(* CODESYS project Simulation_Roboter.project

Project tree, tasks and I/O mapping:
  Device : CODESYS Virtual Control for Linux SL, CODESYS, order no. 2302000005, version 4.22.0.0
    application Application
      libraries: Standard, 3.5.22.0 (System); VisuDialogs, * (System); Unit Conversion Interfaces, * (Intern); CAA Mathematics, * (CAA Technical Workgroup); SM3_Math, * (CODESYS); SysProcess, * (System); CmpBitmapPool, * (System); SysProcess Implementation, * (System)
      task MainTask (cyclic, interval t#20ms, priority 1) calls MAIN_PRG
      task SoftMotion_PlanningTask (cyclic, interval t#2ms, priority 15) calls nothing
      global variables GVL_OPCUA
      visualisation Topics_Vis
      Structs/
        ST_RobotStatus/
          data type ST_RobotStatus
        ST_RobotAction/
          data type ST_RobotAction
          data type Error_Codes_RobotAction
        ST_RobotCommand/
          data type ST_RobotCommand
          data type Status_Codes_RobotCommand
        ST_Orientierung/
          data type ST_euler
          data type ST_quaternions
        ST_Roboter/
          data type ST_Pose_Axis
          data type ST_Pose_TCP
      program MAIN_PRG [FBD]
      FB_Generell/
        function block FB_MoveAction [ST]: MoveToHome, Ex1_ompl_tcp, Ex2_ompl_joint, Ex3_pilz_tcp_ptp, Ex_4_pilz_tcp_lin
        function block FB_Modes [FBD]
        function block FB_RobotStatus [ST]
        function block FB_RobotCommand [ST]
        function block FB_Watchdog [ST]
      program Ablaufkette [SFC]: Ablauf_HomePos, Ablauf_Pos1, Ablauf_Pos2, Ablauf_Pos3, Ablauf_Pos4, Ablauf_Pos5
      Funktionen/
        function FUNC_quat_to_euler [ST]
        function block FB_Quat_to_ZYZ [FBD]
        function block FB_ZYZ_to_Quat [FBD]
        function block FB_Quat_to_ZYX [FBD]
      Symbols
      image pool ImagePool
      visualisation VISU_Auto
      visualisation VISU_Startseite
      visualisation VISU_Manuell
      visualisation VISU_Konfig
      visualisation VISU_Schrittkette
  libraries: SM3_Robotics, * (CODESYS); VisuSymbols, 4.5.0.0 (System)
  text list GlobalTextList
  5ce3da45-db07-42e7-a21c-a00fff4ed8f6|C:\Users\koerp\Documents\Uni\WS2627\04_Projektarbeit-Seitz\Draw_IO\OPC_Strukut.png
  5ce3da45-db07-42e7-a21c-a00fff4ed8f6|C:\Users\koerp\Documents\Uni\WS2627\04_Projektarbeit-Seitz\Draw IO Diagramme\Screenshots\myCobotbeschriftet.png
*)

// Device/Application/Structs/ST_RobotStatus/ST_RobotStatus
// Status Client: Schnittstelle ROS2 <-> SPS
// Ist Zustand des Roboters
TYPE ST_RobotStatus :
STRUCT
	//Ist Gelenkwinkel [rad]
	Ist_Pos_Axis : ST_Pose_Axis; 	
	
	// Ist TCP Pose bezogen auf Roboterbasis
	Ist_Pos_TCP : ST_Pose_TCP;	

	//Verbindungsüberwachung mit Watchdog 
	client_connected : BOOL;
	watchdog_counter : INT;		// Überprüft serverseitige client verbindung
END_STRUCT
END_TYPE

// Device/Application/Structs/ST_RobotCommand/ST_RobotCommand
// Command Client: Schnittstelle ROS2 <-> SPS
// Manuelle Steuerung des Roboters mit MoveIt Servo
TYPE ST_RobotCommand :
STRUCT
	// Gelenke einzeln verfahren
	Mode_Axis: BOOL;					// True: Gelenk Joggen möglich
	Soll_Axis_Servo : ST_Pose_Axis;		//Richtungsvorgabe je Gelenk
	Soll_Axis_Velocity: LREAL;			// Geschwindikeitsvorgabe je Gelenk
	
	// TCP manuell verfahren 
	Mode_TCP: BOOL;						// True: Achsen Joggen möglich
	Soll_TCP_Servo : ST_Pose_TCP;		// Hinweis: Rotation wird nur mit x,y,z übergeben und nicht als Quaternion!
	Soll_TCP_Velocity: LREAL;			// Geschwindkeitsvorgabe für Verfahren
	
	//enable: zum starten und stopen des services servo_node/start_servo und stop_servo
	enable : BOOL;
	
	//Status Code mit Status Codes
	Status_Code: SINT;
	
	// Verbindungsüberwachung mit Watchdog
	client_connected: BOOL;
	watchdog_counter: INT;
END_STRUCT
END_TYPE

// Device/Application/Structs/ST_RobotAction/ST_RobotAction
TYPE ST_RobotAction :
STRUCT
	// Ausführung
	Execute : BOOL;						// TRUE-Puls 
	Error_Code : DINT;					// Ergebnis (int32 MoveItErrorCodes), 1 = SUCCESS,
										// Bedeutung siehe Error_Codes_RobotAction

	// Planer-Auswahl
	Motion_Type : STRING;				// (string pipeline_id) 'ompl' oder 'pilz_industrial_motion_planner'
	Planner_ID : STRING;				// (string planner_id) '' (leer für OMPL), 'PTP' oder 'LIN' für Pilz

	// Art des Ziels (genau eins TRUE)
	Joint_Goal : BOOL;					// TRUE: Gelenkziel -> Soll_Pos_Axis
	TCP_GOAL : BOOL;					// TRUE: kartesisches TCP-Ziel -> Soll_Pos_TCP

	// Planer-Parameter
	num_planning_attempts : DINT;		// (int32 num_planning_attempts) Anzahl Planungsversuche
	allowed_planning_time : LREAL;		// (float64 allowed_planning_time) max. Planungszeit [s]
	max_velocity_scaling : LREAL;		// (float64 max_velocity_scaling_factor) 0..1
	max_acceleration_scaling : LREAL;	// (float64 max_acceleration_scaling_factor) 0..1

	// Zieltoleranzen
	position_tolerance : LREAL;			// (float64) Toleranz TCP-Position [m], gleich für x, y, z
	orientation_tolerance : LREAL;		// (float64) Toleranz TCP-Orientierung [rad], gleich für alle Achsen
	joint_tolerance : LREAL;			// (float64) Toleranz je Gelenk [rad]

	// Zielpose Gelenke [rad]
	Soll_Pos_Axis : ST_Pose_Axis;

	// Zielpose TCP: Position [m], Orientierung als Quaternion
	Soll_Pos_TCP : ST_Pose_TCP;

	// Verbindungsüberwachung mit Watchdog
	client_connected : BOOL;		
	watchdog_counter : INT;				
END_STRUCT
END_TYPE

// Device/Application/Structs/ST_Roboter/ST_Pose_Axis
TYPE ST_Pose_Axis :
STRUCT
	// Gelenkwinkel in rad
	axis_0 : LREAL;
	axis_1 : LREAL;
	axis_2 : LREAL;
	axis_3 : LREAL;
	axis_4 : LREAL;
	axis_5 : LREAL;
END_STRUCT
END_TYPE

// Device/Application/Structs/ST_Roboter/ST_Pose_TCP
TYPE ST_Pose_TCP :
STRUCT
	// Position in m
	trans_x : LREAL;	
	trans_y :  LREAL;
	trans_z : LREAL;
	// Orientierung als Quaternion
	rot_x : LREAL;	// Imaginärteil 	
	rot_y : LREAL;	// Imaginärteil 	
	rot_z : LREAL;	// Imaginärteil 	
	rot_w : LREAL;	//Realteil
END_STRUCT
END_TYPE

// Device/Application/Structs/ST_RobotAction/Error_Codes_RobotAction
{attribute 'qualified_only'}
//{attribute 'strict'}	//CODESYS erlaubt keine TYP Umwandlungen wenn strict aktiv!
{attribute 'to_string'}

TYPE Error_Codes_RobotAction :
(
	NOT_DEFINED := 0,
    SUCCESS := 1,
    FAILURE := 99999,
    PLANNING_FAILED := -1,
    INVALID_MOTION_PLAN := -2,
    MOTION_PLAN_INVALIDATED_BY_ENVIRONMENT_CHANGE := -3,
    CONTROL_FAILED := -4,
    UNABLE_TO_AQUIRE_SENSOR_DATA := -5,
    TIMED_OUT := -6,
    PREEMPTED := -7,
    START_STATE_IN_COLLISION := -10,
    START_STATE_VIOLATES_PATH_CONSTRAINTS := -11,
    START_STATE_INVALID := -26,
    GOAL_IN_COLLISION := -12,
    GOAL_VIOLATES_PATH_CONSTRAINTS := -13,
    GOAL_CONSTRAINTS_VIOLATED := -14,
    GOAL_STATE_INVALID := -27,
    UNRECOGNIZED_GOAL_TYPE := -28,
    INVALID_GROUP_NAME := -15,
    INVALID_GOAL_CONSTRAINTS := -16,
    INVALID_ROBOT_STATE := -17,
    INVALID_LINK_NAME := -18,
    INVALID_OBJECT_NAME := -19,
    FRAME_TRANSFORM_FAILURE := -21,
    COLLISION_CHECKING_UNAVAILABLE := -22,
    ROBOT_STATE_STALE := -23,
    SENSOR_INFO_STALE := -24,
    COMMUNICATION_FAILURE := -25,
    CRASH := -29,
    ABORT := -30,
    NO_IK_SOLUTION := -31
) DINT := NOT_DEFINED;	//Standardwert
END_TYPE

// Device/Application/Structs/ST_Orientierung/ST_euler
//Eulerwinkel intrinsich ZYZ
//ZYZ intrinsisch: bezug auf mitbewegendes Koordinatensystem
//ZYZ extrinsisch: bezug auf festes Koordinatensystem
TYPE ST_euler :
STRUCT
	A : LREAL;	//Z	
	B : LREAL;	//Y
	C : LREAL;	//Z
END_STRUCT
END_TYPE

// Device/Application/Structs/ST_Orientierung/ST_quaternions
TYPE ST_quaternions :
STRUCT
	qx: LREAL;
	qy: LREAL;
	qz: LREAL;
	qw: LREAL;
END_STRUCT
END_TYPE

// Device/Application/Structs/ST_RobotCommand/Status_Codes_RobotCommand
{attribute 'qualified_only'}
//{attribute 'strict'}	//CODESYS erlaubt keine TYP Umwandlungen wenn strict aktiv!
{attribute 'to_string'}
TYPE Status_Codes_RobotCommand :
(
	SERVO_AUS := 99, //wenn Roboter nicht verbunden
	INVALID := -1,
	NO_WARNING := 0,
	DECELERATE_FOR_APPROACHING_SINGULARITY := 1,
	HALT_FOR_SINGULARITY := 2,
	DECELERATE_FOR_LEAVING_SINGULARITY := 3,
	DECELERATE_FOR_COLLISION := 4,
	HALT_FOR_COLLISION := 5,
	JOINT_BOUND := 6	// Achse hat Limit erreich
) SINT := SERVO_AUS;	//Standardwert
END_TYPE

// Device/Application/GVL_OPCUA
{attribute 'qualified_only'}
VAR_GLOBAL
// 	================ Schnittstelle OPC UA =======================================================
	// Schnittstelle Client: ROS2 <-> SPS
	RobotAction: ST_RobotAction;	// Action Client: (Bahnplannung mit MoveIt2)
	RobotStatus : ST_RobotStatus;	// Status Client: Sensorinformationen über Stand des Roboters
	RobotCommand : ST_RobotCommand;	// Command Client: /(Manuelle Steuerung mit MoveIt Servo) 
	// Schnittstelle für SoftKeys 
	// Werden von entrypoint.py Client gelesen, der dann ros2 launch Befehle startet
	Start_RViz2 : BOOL;			//Start RViz2
	Stop_RViz2: BOOL;			//Stop RViz2
	Start_OPCClients: BOOL;		//Start OPC Clients
	Stop_OPC_Clients: BOOL;		//Stop OPC Clients
	
// ================ INTERN ===================================================================	
	Execute : BOOL := FALSE;	//Taster Visu: Ausführen des MoveIt2 Befehls (Auto)
	
	// Ablaufkette
	TIPP : BOOL; 				// Zum Weiterschalten
	Start_Ablaufkette: BOOL;	// Startet Ablaufkette
	Reset_Ablaufkette: BOOL;	//setzt Schrittkette zurück
	
	Joint_Goal : BOOL;			// True: Gelenkziel vorgeben
	TCP_GOAL: BOOL;				// True: Karteisisches TCP Ziel vorgeben
	
	// TCP Sollpositionen (beuogen auf Roboterbasis)
	trans_x : LREAL;	// [m]
	trans_y : LREAL;	// [m]
	trans_z : LREAL;	// [m]
	rot_A : LREAL;		// [°]
	rot_B: LREAL;		// [°]
	rot_C: LREAL;		// [°]
	// Gelenkwinkel Sollpositionen in rad
	axis_0 : LREAL;		// [rad]
	axis_1 : LREAL;		// [rad]
	axis_2 : LREAL;		// [rad]
	axis_3 : LREAL;		// [rad]
	axis_4 : LREAL;		// [rad]
	axis_5 : LREAL;		// [rad]
	// Zieltoleranzen
	position_tolerance : LREAL;			// Toleranz TCP Position [m]
	orientation_tolerance : LREAL;		// Toleranz TCP Orientierung [rad]
	joint_tolerance: LREAL;				// Tolerant Achswinkel in [rad]

	Motion_Type : STRING;				// pipeline_id: "ompl" oder "pilz_industrial_motion_planner"
	Planner_ID : STRING;				// planner_id: " " (leer für OMPL) "PTP" oder "LIN" für Pilz

	num_planning_attempts : DINT;		// Anzahl Plannungsversuche
	allowed_planning_time : LREAL;		// max Plannungszeit in s
	max_velocity_scaling : LREAL;		// 0 .. 1 Skalierung maximale Gelenkgeschwindigkeit
	max_acceleration_scaling : LREAL;	// 0 ...1 Skalierung maximale Gelenkbeschleunigung
END_VAR

VAR_GLOBAL CONSTANT
	PI : REAL := 3.14159;
END_VAR

// Device/Application/MAIN_PRG
PROGRAM MAIN_PRG
VAR
// ======== Betriebsart ==============================================================
	Modes : FB_Modes;						// Auswahl Hand / Automatik (Hand hat Vorrang)
	
// ========Automatik ==============================================================
	// Automatik: Bewegungsauftrag an MoveIt 2 (Action Client)
	RobotAction : FB_MoveAction;			// Übergibt Sollwerte aus GVL_OPCUA an RobotAction
	trig : R_TRIG;							// Flanke von GVL_OPCUA.Execute 
	Action_zyz_to_quat : FB_ZYZ_to_Quat;	// Soll-Orientierung ZYZ -> Quaternion
	Status_Error_Codes_Action : Error_Codes_RobotAction;	// Ergebnis der Bewegung 

	// Vorgefertigte Beispielbewegungen 
	xMoveHome : BOOL;						
	xEx1_ompl_tcp : BOOL;				
	xEx2_ompl_joint : BOOL;				
	xEx3_pilz_tcp_ptp : BOOL;			
	xEx4_pilz_tcp_lin : BOOL;			

// ============Handbetrieb ==========================================================
	// Handbetrieb: Joggen über MoveIt Servo (Command Client)

	RobotCommand : FB_RobotCommand;		
	Status_Servo : Status_Codes_RobotCommand;	// Statuscode MoveIt Servo 

// ==============Istwerte========================================================
	// Istwerte und Verbindungsüberwachung (Status Client)
	RobotStatus : FB_RobotStatus;			// Watchdog Status Client
	Status_Quat_to_ZYZ : FB_Quat_to_ZYZ;	// Ist-Orientierung TCP Quaternion -> ZYZ 
END_VAR

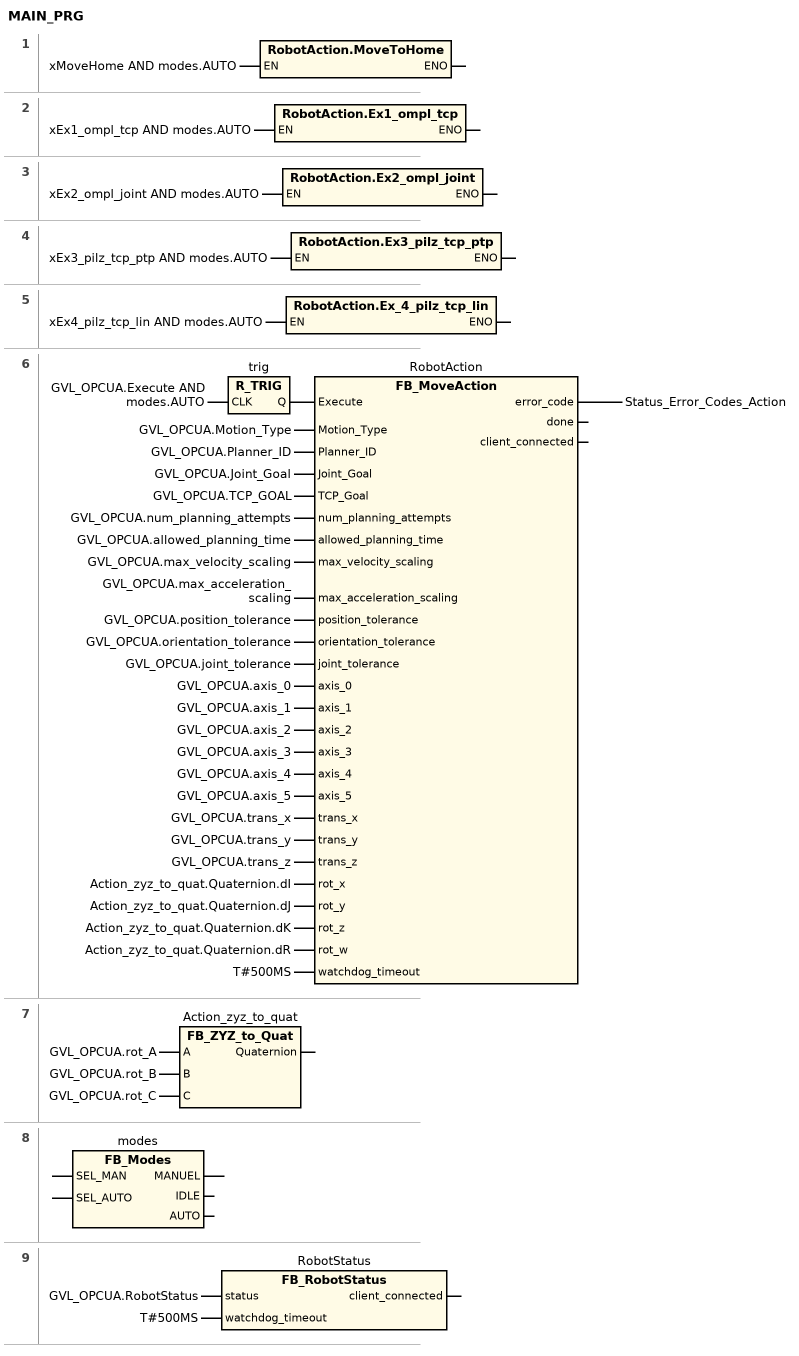
// NETWORK 1
IF xMoveHome AND modes.AUTO THEN RobotAction.MoveToHome(); END_IF

// NETWORK 2
IF xEx1_ompl_tcp AND modes.AUTO THEN RobotAction.Ex1_ompl_tcp(); END_IF

// NETWORK 3
IF xEx2_ompl_joint AND modes.AUTO THEN RobotAction.Ex2_ompl_joint(); END_IF

// NETWORK 4
IF xEx3_pilz_tcp_ptp AND modes.AUTO THEN RobotAction.Ex3_pilz_tcp_ptp(); END_IF

// NETWORK 5
IF xEx4_pilz_tcp_lin AND modes.AUTO THEN RobotAction.Ex_4_pilz_tcp_lin(); END_IF

// NETWORK 6
trig(CLK := GVL_OPCUA.Execute AND modes.AUTO); // R_TRIG
RobotAction(
    Execute := trig.Q,
    Motion_Type := GVL_OPCUA.Motion_Type,
    Planner_ID := GVL_OPCUA.Planner_ID,
    Joint_Goal := GVL_OPCUA.Joint_Goal,
    TCP_Goal := GVL_OPCUA.TCP_GOAL,
    num_planning_attempts := GVL_OPCUA.num_planning_attempts,
    allowed_planning_time := GVL_OPCUA.allowed_planning_time,
    max_velocity_scaling := GVL_OPCUA.max_velocity_scaling,
    max_acceleration_scaling := GVL_OPCUA.max_acceleration_scaling,
    position_tolerance := GVL_OPCUA.position_tolerance,
    orientation_tolerance := GVL_OPCUA.orientation_tolerance,
    joint_tolerance := GVL_OPCUA.joint_tolerance,
    axis_0 := GVL_OPCUA.axis_0,
    axis_1 := GVL_OPCUA.axis_1,
    axis_2 := GVL_OPCUA.axis_2,
    axis_3 := GVL_OPCUA.axis_3,
    axis_4 := GVL_OPCUA.axis_4,
    axis_5 := GVL_OPCUA.axis_5,
    trans_x := GVL_OPCUA.trans_x,
    trans_y := GVL_OPCUA.trans_y,
    trans_z := GVL_OPCUA.trans_z,
    rot_x := Action_zyz_to_quat.Quaternion.dI,
    rot_y := Action_zyz_to_quat.Quaternion.dJ,
    rot_z := Action_zyz_to_quat.Quaternion.dK,
    rot_w := Action_zyz_to_quat.Quaternion.dR,
    watchdog_timeout := T#500MS); // FB_MoveAction
Status_Error_Codes_Action := RobotAction.error_code;

// NETWORK 7
Action_zyz_to_quat(A := GVL_OPCUA.rot_A, B := GVL_OPCUA.rot_B, C := GVL_OPCUA.rot_C); // FB_ZYZ_to_Quat

// NETWORK 8
modes(); // FB_Modes

// NETWORK 9
RobotStatus(status := GVL_OPCUA.RobotStatus, watchdog_timeout := T#500MS); // FB_RobotStatus

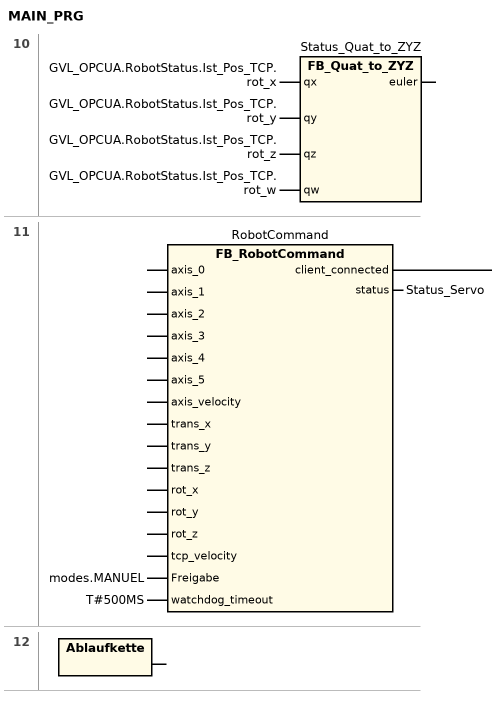
// NETWORK 10
Status_Quat_to_ZYZ(
    qx := GVL_OPCUA.RobotStatus.Ist_Pos_TCP.rot_x,
    qy := GVL_OPCUA.RobotStatus.Ist_Pos_TCP.rot_y,
    qz := GVL_OPCUA.RobotStatus.Ist_Pos_TCP.rot_z,
    qw := GVL_OPCUA.RobotStatus.Ist_Pos_TCP.rot_w); // FB_Quat_to_ZYZ

// NETWORK 11
RobotCommand(Freigabe := modes.MANUEL, watchdog_timeout := T#500MS, status => Status_Servo); // FB_RobotCommand

// NETWORK 12
Ablaufkette();

END_PROGRAM

// Device/Application/FB_Generell/FB_MoveAction
FUNCTION_BLOCK FB_MoveAction
// Übergabe von Gelenk oder ZCP Ziel an ROS2 Client
VAR_INPUT
    Execute : BOOL;

    Motion_Type : STRING;
    Planner_ID : STRING;

    Joint_Goal : BOOL;
    TCP_Goal : BOOL;

    num_planning_attempts : DINT;
    allowed_planning_time : LREAL;

    max_velocity_scaling : LREAL;
    max_acceleration_scaling : LREAL;

    position_tolerance : LREAL;
    orientation_tolerance : LREAL;
	joint_tolerance: LREAL;

    // Joints
    axis_0 : LREAL;
    axis_1 : LREAL;
    axis_2 : LREAL;
    axis_3 : LREAL;
    axis_4 : LREAL;
    axis_5 : LREAL;

    // TCP
    trans_x : LREAL;
    trans_y : LREAL;
    trans_z : LREAL;
    rot_x : LREAL;
    rot_y : LREAL;
    rot_z : LREAL;
    rot_w : LREAL;
	
	watchdog_timeout : TIME := T#500MS;	//Timeout des Watchdogs
END_VAR
VAR_OUTPUT
	error_code:DINT;
	done : BOOL;
	//Watchdog
	client_connected : BOOL;
END_VAR
VAR
	watchdog : FB_Watchdog;
END_VAR

//Watchdog aktualisieren
watchdog(watchdog_counter := GVL_OPCUA.RobotAction.watchdog_counter, timeout := watchdog_timeout);
client_connected := watchdog.client_connected;

// Execute
GVL_OPCUA.RobotAction.Execute := Execute;

// Allgemein
GVL_OPCUA.RobotAction.Motion_Type := Motion_Type;
GVL_OPCUA.RobotAction.Planner_ID := Planner_ID;

GVL_OPCUA.RobotAction.Joint_Goal := Joint_Goal;
GVL_OPCUA.RobotAction.TCP_GOAL := TCP_Goal;

GVL_OPCUA.RobotAction.num_planning_attempts := num_planning_attempts;
GVL_OPCUA.RobotAction.allowed_planning_time := allowed_planning_time;

GVL_OPCUA.RobotAction.max_velocity_scaling := max_velocity_scaling;
GVL_OPCUA.RobotAction.max_acceleration_scaling := max_acceleration_scaling;

GVL_OPCUA.RobotAction.position_tolerance := position_tolerance;
GVL_OPCUA.RobotAction.orientation_tolerance := orientation_tolerance;
GVL_OPCUA.RobotAction.joint_tolerance := joint_tolerance;

// Joints
GVL_OPCUA.RobotAction.Soll_Pos_Axis.axis_0 := axis_0;
GVL_OPCUA.RobotAction.Soll_Pos_Axis.axis_1 := axis_1;
GVL_OPCUA.RobotAction.Soll_Pos_Axis.axis_2 := axis_2;
GVL_OPCUA.RobotAction.Soll_Pos_Axis.axis_3 := axis_3;
GVL_OPCUA.RobotAction.Soll_Pos_Axis.axis_4 := axis_4;
GVL_OPCUA.RobotAction.Soll_Pos_Axis.axis_5 := axis_5;


// TCP
GVL_OPCUA.RobotAction.Soll_Pos_TCP.trans_x := trans_x;
GVL_OPCUA.RobotAction.Soll_Pos_TCP.trans_y := trans_y;
GVL_OPCUA.RobotAction.Soll_Pos_TCP.trans_z := trans_z;

GVL_OPCUA.RobotAction.Soll_Pos_TCP.rot_x := rot_x;
GVL_OPCUA.RobotAction.Soll_Pos_TCP.rot_y := rot_y;
GVL_OPCUA.RobotAction.Soll_Pos_TCP.rot_z := rot_z;
GVL_OPCUA.RobotAction.Soll_Pos_TCP.rot_w := rot_w;

//OUTPUT
error_code := GVL_OPCUA.RobotAction.Error_Code;
IF error_code = 1 THEN
	done := TRUE;
ELSE 
	done := FALSE;
END_IF

ACTION MoveToHome:
//HomePosition
GVL_OPCUA.Joint_Goal := TRUE;
GVL_OPCUA.TCP_Goal := FALSE;

GVL_OPCUA.axis_0 := 0.0;
GVL_OPCUA.axis_1 := 0.0;
GVL_OPCUA.axis_2 := 0.0;
GVL_OPCUA.axis_3 := 0.0;
GVL_OPCUA.axis_4 := 0.0;
GVL_OPCUA.axis_5 := 0.0;

GVL_OPCUA.joint_tolerance := 0.005;

GVL_OPCUA.Motion_Type := 'ompl';
GVL_OPCUA.Planner_ID := '';

GVL_OPCUA.num_planning_attempts := 5;
GVL_OPCUA.allowed_planning_time := 5;
GVL_OPCUA.max_velocity_scaling := 0.1;
GVL_OPCUA.max_acceleration_scaling := 0.1;
END_ACTION

ACTION Ex1_ompl_tcp:
GVL_OPCUA.Joint_Goal := FALSE;
GVL_OPCUA.TCP_Goal := TRUE;

GVL_OPCUA.trans_x := 0.114;
GVL_OPCUA.trans_y := -0.019;
GVL_OPCUA.trans_z := 0.357;
GVL_OPCUA.rot_A := 0.0;
GVL_OPCUA.rot_B := 90.0;
GVL_OPCUA.rot_C := -90.0;

GVL_OPCUA.position_tolerance := 0.02;
GVL_OPCUA.orientation_tolerance := 0.05;

GVL_OPCUA.Motion_Type := 'ompl';
GVL_OPCUA.Planner_ID := '';

GVL_OPCUA.num_planning_attempts := 5;
GVL_OPCUA.allowed_planning_time := 5;
GVL_OPCUA.max_velocity_scaling := 0.2;
GVL_OPCUA.max_acceleration_scaling := 0.2;
END_ACTION

ACTION Ex2_ompl_joint:
GVL_OPCUA.Joint_Goal := TRUE;
GVL_OPCUA.TCP_Goal := FALSE;

GVL_OPCUA.axis_0 := 0.1;
GVL_OPCUA.axis_1 := -1.65;
GVL_OPCUA.axis_2 := 1.7;
GVL_OPCUA.axis_3 := 0.1;
GVL_OPCUA.axis_4 := 0.2;
GVL_OPCUA.axis_5 := 0.3;

GVL_OPCUA.Motion_Type := 'ompl';
GVL_OPCUA.Planner_ID := '';

GVL_OPCUA.joint_tolerance := 0.01;

GVL_OPCUA.num_planning_attempts := 5;
GVL_OPCUA.allowed_planning_time := 5;
GVL_OPCUA.max_velocity_scaling := 0.2;
GVL_OPCUA.max_acceleration_scaling := 0.2;
END_ACTION

ACTION Ex3_pilz_tcp_ptp:
GVL_OPCUA.Joint_Goal := FALSE;
GVL_OPCUA.TCP_Goal := TRUE;

GVL_OPCUA.trans_x := 0.17;
GVL_OPCUA.trans_y := -0.04;
GVL_OPCUA.trans_z := 0.22;
GVL_OPCUA.rot_A := 0.0;
GVL_OPCUA.rot_B := 90.0;
GVL_OPCUA.rot_C := -90.0;

GVL_OPCUA.position_tolerance := 0.02;
GVL_OPCUA.orientation_tolerance := 0.05;

GVL_OPCUA.Motion_Type := 'pilz_industrial_motion_planner';
GVL_OPCUA.Planner_ID := 'PTP';

GVL_OPCUA.num_planning_attempts := 10;
GVL_OPCUA.allowed_planning_time := 10;
GVL_OPCUA.max_velocity_scaling := 0.05;
GVL_OPCUA.max_acceleration_scaling := 0.05;
END_ACTION

ACTION Ex_4_pilz_tcp_lin:
GVL_OPCUA.Joint_Goal := FALSE;
GVL_OPCUA.TCP_Goal := TRUE;

GVL_OPCUA.trans_x := 0.2;
GVL_OPCUA.trans_y := -0.041;
GVL_OPCUA.trans_z := 0.3;
GVL_OPCUA.rot_A := 0.0;
GVL_OPCUA.rot_B := 90.0;
GVL_OPCUA.rot_C := -90.0;

GVL_OPCUA.Motion_Type := 'pilz_industrial_motion_planner';
GVL_OPCUA.Planner_ID := 'LIN';

GVL_OPCUA.position_tolerance := 0.02;
GVL_OPCUA.orientation_tolerance := 0.05;

GVL_OPCUA.num_planning_attempts := 10;
GVL_OPCUA.allowed_planning_time := 10;
GVL_OPCUA.max_velocity_scaling := 0.005;
GVL_OPCUA.max_acceleration_scaling := 0.005;
END_ACTION

END_FUNCTION_BLOCK

// Device/Application/FB_Generell/FB_Watchdog
FUNCTION_BLOCK FB_Watchdog
VAR_INPUT
	Watchdog_counter: INT;	// Zähler im ROS2 Programm
	Timeout : TIME := T#500MS;
END_VAR
VAR
	//Watchdog
	Watchdog_counter_old : INT := 0;
	Timer : TON;
END_VAR
VAR_OUTPUT
	client_connected: BOOL;	//Anzeige ob verbunden
END_VAR

//Watchdog zum Testen ob noch mit Client verbunden!
IF Watchdog_counter <> Watchdog_counter_old THEN
	Watchdog_counter_old :=  Watchdog_counter;
    client_connected := TRUE;
    Timer(IN := FALSE);
ELSE
    Timer(IN := TRUE,PT := Timeout );
END_IF;
IF Timer.Q THEN
    client_connected := FALSE;
END_IF;

END_FUNCTION_BLOCK

// Device/Application/Funktionen/FB_ZYZ_to_Quat
FUNCTION_BLOCK FB_ZYZ_to_Quat
VAR_INPUT
	A : LREAL;
	B: LREAL;
	C: LREAL;
END_VAR
VAR_OUTPUT
	Quaternion: SMC_Quat;
END_VAR
VAR
	Rotation_Matrix: SMC_Matrix3;
END_VAR

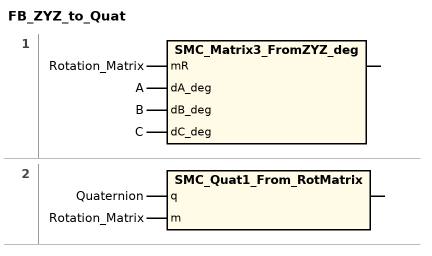
// NETWORK 1
SMC_Matrix3_FromZYZ_deg(mR := Rotation_Matrix, dA_deg := A, dB_deg := B, dC_deg := C);

// NETWORK 2
SMC_Quat1_From_RotMatrix(q := Quaternion, m := Rotation_Matrix);

END_FUNCTION_BLOCK

// Device/Application/FB_Generell/FB_Modes
FUNCTION_BLOCK FB_Modes	// Betriebsartenumschaltung mit Betriebsartenhierachie MAN > AUTO
VAR_INPUT
	SEL_MAN : BOOL;
	SEL_AUTO: BOOL;
END_VAR
VAR_OUTPUT
	MANUEL : BOOL;	//z1
	IDLE: BOOL;		//z0
	AUTO: BOOL;		//z2
END_VAR
VAR
	z0, z1, z2 : BOOL;
	H1, H2: RS;
	z: INT;
END_VAR
VAR // added by the converter: edge detectors and wires of the graphical bodies
    _w1, _w2, _w3 : BOOL;
END_VAR

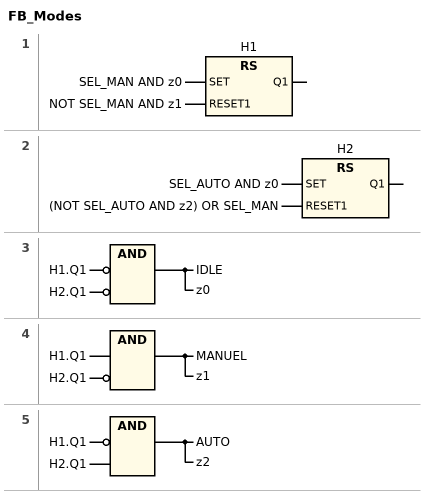
// NETWORK 1
H1(SET := SEL_MAN AND z0, RESET1 := NOT SEL_MAN AND z1); // RS

// NETWORK 2
H2(SET := SEL_AUTO AND z0, RESET1 := (NOT SEL_AUTO AND z2) OR SEL_MAN); // RS

// NETWORK 3
_w1 := NOT H1.Q1 AND NOT H2.Q1;
IDLE := _w1;
z0 := _w1;

// NETWORK 4
_w2 := H1.Q1 AND NOT H2.Q1;
MANUEL := _w2;
z1 := _w2;

// NETWORK 5
_w3 := NOT H1.Q1 AND H2.Q1;
AUTO := _w3;
z2 := _w3;

END_FUNCTION_BLOCK

// Device/Application/FB_Generell/FB_RobotStatus
FUNCTION_BLOCK FB_RobotStatus
VAR_INPUT
	status: ST_RobotStatus;
	watchdog_timeout: TIME := T#500MS;
END_VAR
VAR_OUTPUT
	client_connected : BOOL;
END_VAR
VAR
	watchdog : FB_Watchdog;
END_VAR

//Watchdog aktualisieren
watchdog(watchdog_counter := status.watchdog_counter, timeout := watchdog_timeout);
client_connected := watchdog.client_connected;

END_FUNCTION_BLOCK

// Device/Application/Funktionen/FB_Quat_to_ZYZ
FUNCTION_BLOCK FB_Quat_to_ZYZ
VAR_INPUT
	qx : LREAL;
	qy: LREAL;
	qz:LREAL;
	qw : LREAL;

END_VAR
VAR_OUTPUT
	euler : ST_euler;
END_VAR
VAR
	Quaternion: SMC_Quat;
	Rotation_Matrix: SMC_Matrix3;
END_VAR

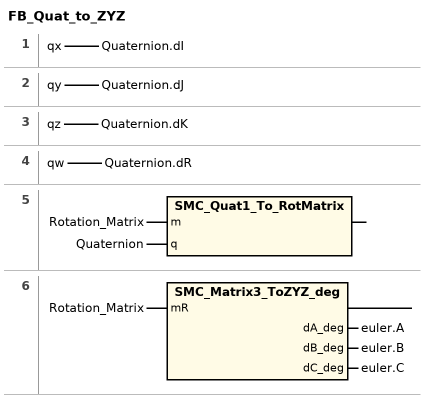
// NETWORK 1
Quaternion.dI := qx;

// NETWORK 2
Quaternion.dJ := qy;

// NETWORK 3
Quaternion.dK := qz;

// NETWORK 4
Quaternion.dR := qw;

// NETWORK 5
SMC_Quat1_To_RotMatrix(m := Rotation_Matrix, q := Quaternion);

// NETWORK 6
SMC_Matrix3_ToZYZ_deg(mR := Rotation_Matrix, dA_deg => euler.A, dB_deg => euler.B, dC_deg => euler.C);

END_FUNCTION_BLOCK

// Device/Application/FB_Generell/FB_RobotCommand
FUNCTION_BLOCK FB_RobotCommand
VAR_INPUT
	axis_0 : LREAL;
	axis_1 : LREAL;
	axis_2: LREAL;
	axis_3 : LREAL;
	axis_4 : LREAL;
	axis_5 : LREAL;
	axis_velocity : LREAL;
	
	trans_x : LREAL;
	trans_y : LREAL;
	trans_z : LREAL;
	rot_x : LREAL;
	rot_y : LREAL;
	rot_z : LREAL;
	tcp_velocity : LREAL;
	
	//Allgemein
	Freigabe:BOOL:=FALSE;
	
	watchdog_timeout: TIME := T#500MS;
END_VAR
VAR_OUTPUT
	// Watchdog
	client_connected : BOOL;
	// Status Meldung
	status: SINT;	//Datentyp INT8
END_VAR
VAR
	//Watchdog
	watchdog : FB_Watchdog;
END_VAR

//Watchdog aktualisieren
watchdog(watchdog_counter := GVL_OPCUA.RobotCommand.watchdog_counter, timeout := watchdog_timeout);
client_connected := watchdog.client_connected;

IF Freigabe THEN	//Freigabe wenn manueller Betrieb
	GVL_OPCUA.RobotCommand.Soll_Axis_Servo.axis_0 := axis_0;
	GVL_OPCUA.RobotCommand.Soll_Axis_Servo.axis_1 := axis_1;
	GVL_OPCUA.RobotCommand.Soll_Axis_Servo.axis_2 := axis_2;
	GVL_OPCUA.RobotCommand.Soll_Axis_Servo.axis_3 := axis_3;
	GVL_OPCUA.RobotCommand.Soll_Axis_Servo.axis_4 := axis_4;
	GVL_OPCUA.RobotCommand.Soll_Axis_Servo.axis_5 := axis_5;
	GVL_OPCUA.RobotCommand.Soll_Axis_Velocity := axis_velocity;
	
	GVL_OPCUA.RobotCommand.Soll_TCP_Servo.trans_x := trans_x;
	GVL_OPCUA.RobotCommand.Soll_TCP_Servo.trans_y := trans_y;
	GVL_OPCUA.RobotCommand.Soll_TCP_Servo.trans_z := trans_z;
	GVL_OPCUA.RobotCommand.Soll_TCP_Servo.rot_x := rot_x;
	GVL_OPCUA.RobotCommand.Soll_TCP_Servo.rot_y := rot_y;
	GVL_OPCUA.RobotCommand.Soll_TCP_Servo.rot_z := rot_z;
	GVL_OPCUA.RobotCommand.Soll_TCP_Velocity := tcp_velocity;
	
	// start der /servo_node/start_servo
	GVL_OPCUA.RobotCommand.enable := TRUE;
	
ELSE
	GVL_OPCUA.RobotCommand.enable := FALSE;
END_IF

// Status Code
status := GVL_OPCUA.RobotCommand.Status_Code;

END_FUNCTION_BLOCK

// Device/Application/Ablaufkette
PROGRAM Ablaufkette
VAR
	SFCCurrentStep : STRING;
END_VAR

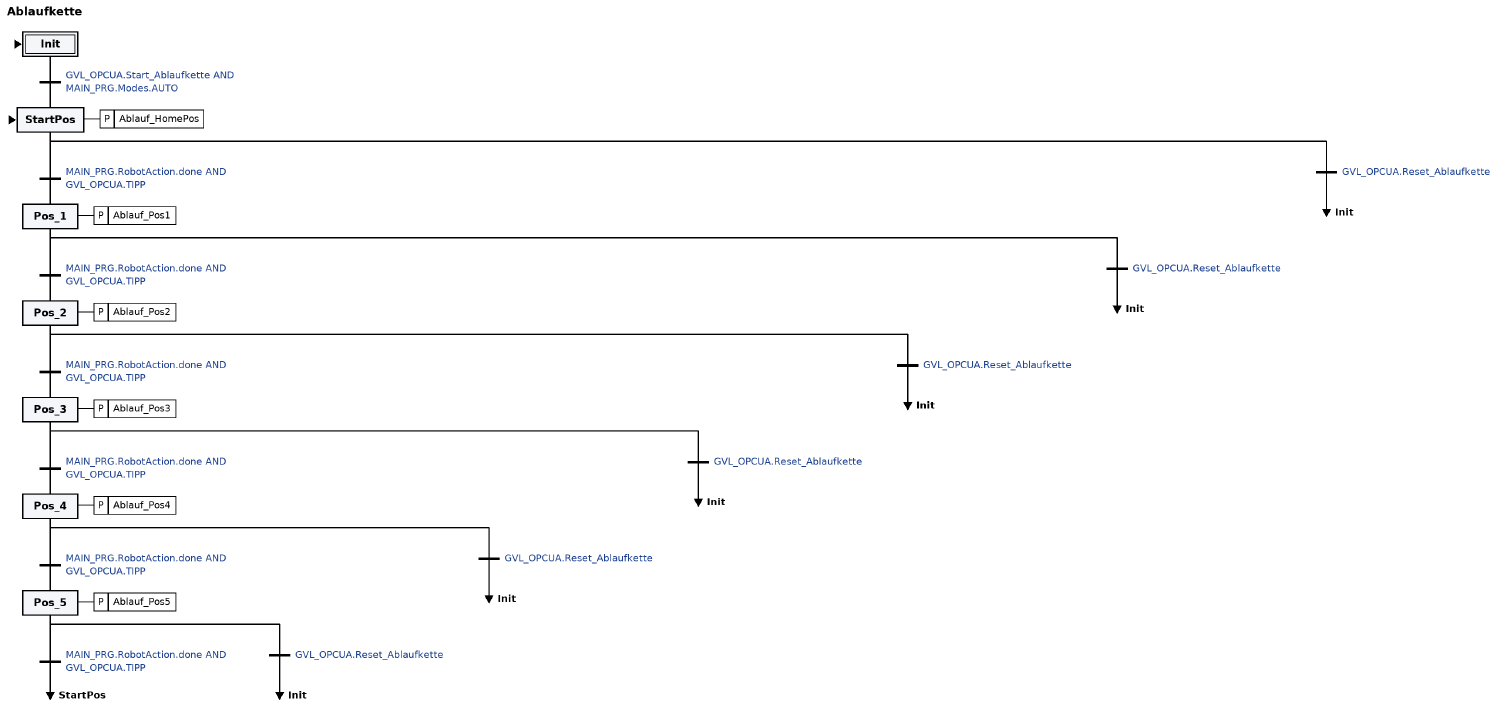
INITIAL_STEP Init:
END_STEP
TRANSITION FROM Init TO StartPos
    := GVL_OPCUA.Start_Ablaufkette AND MAIN_PRG.Modes.AUTO;
END_TRANSITION
STEP StartPos:  // min time t#1s
    Ablauf_HomePos(P);
END_STEP
TRANSITION FROM StartPos TO Pos_1
    := MAIN_PRG.RobotAction.done AND GVL_OPCUA.TIPP;
END_TRANSITION
TRANSITION FROM StartPos TO Init
    := GVL_OPCUA.Reset_Ablaufkette;
END_TRANSITION
STEP Pos_1:  // min time t#1s
    Ablauf_Pos1(P);
END_STEP
TRANSITION FROM Pos_1 TO Pos_2
    := MAIN_PRG.RobotAction.done AND GVL_OPCUA.TIPP;
END_TRANSITION
TRANSITION FROM Pos_1 TO Init
    := GVL_OPCUA.Reset_Ablaufkette;
END_TRANSITION
STEP Pos_2:  // min time t#1s
    Ablauf_Pos2(P);
END_STEP
TRANSITION FROM Pos_2 TO Pos_3
    := MAIN_PRG.RobotAction.done AND GVL_OPCUA.TIPP;
END_TRANSITION
TRANSITION FROM Pos_2 TO Init
    := GVL_OPCUA.Reset_Ablaufkette;
END_TRANSITION
STEP Pos_3:  // min time t#1s
    Ablauf_Pos3(P);
END_STEP
TRANSITION FROM Pos_3 TO Pos_4
    := MAIN_PRG.RobotAction.done AND GVL_OPCUA.TIPP;
END_TRANSITION
TRANSITION FROM Pos_3 TO Init
    := GVL_OPCUA.Reset_Ablaufkette;
END_TRANSITION
STEP Pos_4:  // min time t#1s
    Ablauf_Pos4(P);
END_STEP
TRANSITION FROM Pos_4 TO Pos_5
    := MAIN_PRG.RobotAction.done AND GVL_OPCUA.TIPP;
END_TRANSITION
TRANSITION FROM Pos_4 TO Init
    := GVL_OPCUA.Reset_Ablaufkette;
END_TRANSITION
STEP Pos_5:  // min time t#1s
    Ablauf_Pos5(P);
END_STEP
TRANSITION FROM Pos_5 TO StartPos
    := MAIN_PRG.RobotAction.done AND GVL_OPCUA.TIPP;
END_TRANSITION
TRANSITION FROM Pos_5 TO Init
    := GVL_OPCUA.Reset_Ablaufkette;
END_TRANSITION

ACTION Ablauf_HomePos:
GVL_OPCUA.Joint_Goal := TRUE;
GVL_OPCUA.TCP_Goal := FALSE;

GVL_OPCUA.axis_0 := 0.10;
GVL_OPCUA.axis_1 := -0.1;
GVL_OPCUA.axis_2 := -1.6;
GVL_OPCUA.axis_3 := 1.7;
GVL_OPCUA.axis_4 := 0.1;
GVL_OPCUA.axis_5 := 0.2;

GVL_OPCUA.joint_tolerance := 0.01;

GVL_OPCUA.Motion_Type := 'ompl';
GVL_OPCUA.Planner_ID := '';

GVL_OPCUA.num_planning_attempts := 10;
GVL_OPCUA.allowed_planning_time := 10;

GVL_OPCUA.max_velocity_scaling := 0.2;
GVL_OPCUA.max_acceleration_scaling := 0.2;
END_ACTION

ACTION Ablauf_Pos1:
GVL_OPCUA.Joint_Goal := FALSE;
GVL_OPCUA.TCP_Goal := TRUE;

GVL_OPCUA.trans_x := 0.18;
GVL_OPCUA.trans_y := -0.0;
GVL_OPCUA.trans_z := 0.3;

GVL_OPCUA.rot_A := 0.0;
GVL_OPCUA.rot_B := 90.0;
GVL_OPCUA.rot_C := -90.0;

GVL_OPCUA.position_tolerance := 0.005;
GVL_OPCUA.orientation_tolerance := 0.05;

GVL_OPCUA.Motion_Type := 'ompl';
GVL_OPCUA.Planner_ID := '';

GVL_OPCUA.num_planning_attempts := 10;
GVL_OPCUA.allowed_planning_time := 10;
GVL_OPCUA.max_velocity_scaling := 0.1;
GVL_OPCUA.max_acceleration_scaling := 0.1;
END_ACTION

ACTION Ablauf_Pos2:
GVL_OPCUA.Joint_Goal := FALSE;
GVL_OPCUA.TCP_Goal := TRUE;

GVL_OPCUA.trans_x := 0.18;
GVL_OPCUA.trans_y := 0.05;
GVL_OPCUA.trans_z := 0.3;

GVL_OPCUA.rot_A := 0.0;
GVL_OPCUA.rot_B := 90.0;
GVL_OPCUA.rot_C := -90.0;

GVL_OPCUA.position_tolerance := 0.005;
GVL_OPCUA.orientation_tolerance := 0.05;

GVL_OPCUA.Motion_Type := 'pilz_industrial_motion_planner';
GVL_OPCUA.Planner_ID := 'PTP';

GVL_OPCUA.num_planning_attempts := 10;
GVL_OPCUA.allowed_planning_time := 10;
GVL_OPCUA.max_velocity_scaling := 0.1;
GVL_OPCUA.max_acceleration_scaling := 0.1;
END_ACTION

ACTION Ablauf_Pos3:
GVL_OPCUA.Joint_Goal := FALSE;
GVL_OPCUA.TCP_Goal := TRUE;

GVL_OPCUA.trans_x := 0.18;
GVL_OPCUA.trans_y := 0.05;
GVL_OPCUA.trans_z := 0.2;

GVL_OPCUA.rot_A := 0.0;
GVL_OPCUA.rot_B := 90.0;
GVL_OPCUA.rot_C := -90.0;

GVL_OPCUA.position_tolerance := 0.005;
GVL_OPCUA.orientation_tolerance := 0.05;

GVL_OPCUA.Motion_Type := 'pilz_industrial_motion_planner';
GVL_OPCUA.Planner_ID := 'PTP';

GVL_OPCUA.num_planning_attempts := 10;
GVL_OPCUA.allowed_planning_time := 10;
GVL_OPCUA.max_velocity_scaling := 0.1;
GVL_OPCUA.max_acceleration_scaling := 0.1;
END_ACTION

ACTION Ablauf_Pos4:
GVL_OPCUA.Joint_Goal := FALSE;
GVL_OPCUA.TCP_Goal := TRUE;

GVL_OPCUA.trans_x := 0.18;
GVL_OPCUA.trans_y := -0.05;
GVL_OPCUA.trans_z := 0.2;

GVL_OPCUA.rot_A := 0.0;
GVL_OPCUA.rot_B := 90.0;
GVL_OPCUA.rot_C := -90.0;

GVL_OPCUA.position_tolerance := 0.005;
GVL_OPCUA.orientation_tolerance := 0.05;

GVL_OPCUA.Motion_Type := 'pilz_industrial_motion_planner';
GVL_OPCUA.Planner_ID := 'PTP';

GVL_OPCUA.num_planning_attempts := 10;
GVL_OPCUA.allowed_planning_time := 10;
GVL_OPCUA.max_velocity_scaling := 0.1;
GVL_OPCUA.max_acceleration_scaling := 0.1;
END_ACTION

ACTION Ablauf_Pos5:
GVL_OPCUA.Joint_Goal := FALSE;
GVL_OPCUA.TCP_Goal := TRUE;

GVL_OPCUA.trans_x := 0.18;
GVL_OPCUA.trans_y := -0.05;
GVL_OPCUA.trans_z := 0.3;

GVL_OPCUA.rot_A := 0.0;
GVL_OPCUA.rot_B := 90.0;
GVL_OPCUA.rot_C := -90.0;

GVL_OPCUA.position_tolerance := 0.005;
GVL_OPCUA.orientation_tolerance := 0.05;

GVL_OPCUA.Motion_Type := 'pilz_industrial_motion_planner';
GVL_OPCUA.Planner_ID := 'PTP';

GVL_OPCUA.num_planning_attempts := 10;
GVL_OPCUA.allowed_planning_time := 10;
GVL_OPCUA.max_velocity_scaling := 0.1;
GVL_OPCUA.max_acceleration_scaling := 0.1;
END_ACTION

END_PROGRAM

// Device/Application/Funktionen/FUNC_quat_to_euler
FUNCTION FUNC_quat_to_euler : ST_euler
VAR_INPUT
	qx : LREAL;
	qy : LREAL;
	qz : LREAL;
	qw : LREAL;
END_VAR
VAR
	r11, r12, r13, r21, r22, r23, r31, r32, r33 : LREAL;
	const_epsilon : LREAL := 1.0E-6; // Toleranz für Gimbal Lock
	result : ST_euler;
	
END_VAR

//Quaternion -> Euler mit ZYZ (intrinsisch) 
//Ausgabe der Euler Winkel in Grad
//Rotationsmatrix Quaternion
r11 := 1.0 - 2.0 * (qy*qy + qz*qz);
r12 := 2.0 * (qx*qy - qz*qw);
r13 := 2.0 * (qx*qz + qy*qw);

r21 := 2.0 * (qx*qy + qz*qw);
r22 := 1.0 - 2.0 * (qx*qx + qz*qz);
r23 := 2.0 * (qy*qz - qx*qw);

r31 := 2.0 * (qx*qz - qy*qw);
r32 := 2.0 * (qy*qz + qx*qw);
r33 := 1.0 - 2.0 * (qx*qx + qy*qy);

result.B := MATH.atan2_func(SQRT(r31*r31+r32*r32),r33);

IF result.B < const_epsilon THEN
	//Gimbal Lock Nordpol
	result.A := 0.0;
	result.C := MATH.atan2_func(r21,r11);
	
ELSIF result.B > (MATH.PI - const_epsilon) THEN
	//Gimbal Lock Südpol
	result.A := 0.0;
	result.C := MATH.atan2_func(-r21,-r11);
ELSE
	//normal
	result.A := MATH.atan2_func(r23,r13);
	result.C := MATH.atan2_func(r32,-r31);
	
END_IF

result.A := result.A * (180.0/MATH.PI);
result.B := result.B * (180.0/MATH.PI);
result.C := result.C * (180.0/MATH.PI);

FUNC_quat_to_euler := result;

END_FUNCTION

// Device/Application/Funktionen/FB_Quat_to_ZYX
FUNCTION_BLOCK FB_Quat_to_ZYX
VAR_INPUT
	qx : LREAL;
	qy: LREAL;
	qz:LREAL;
	qw : LREAL;

END_VAR
VAR_OUTPUT
	euler : ST_euler;
END_VAR
VAR
	Quaternion: SMC_Quat;
	Rotation_Matrix: SMC_Matrix3;
END_VAR

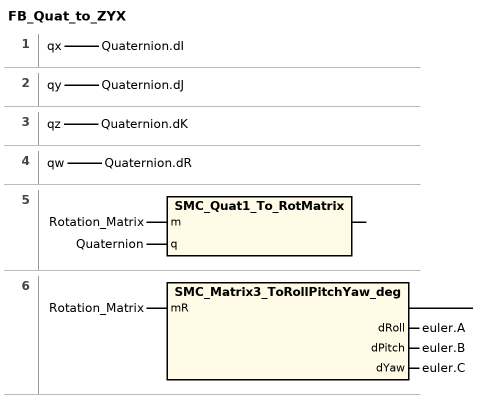
// NETWORK 1
Quaternion.dI := qx;

// NETWORK 2
Quaternion.dJ := qy;

// NETWORK 3
Quaternion.dK := qz;

// NETWORK 4
Quaternion.dR := qw;

// NETWORK 5
SMC_Quat1_To_RotMatrix(m := Rotation_Matrix, q := Quaternion);

// NETWORK 6
SMC_Matrix3_ToRollPitchYaw_deg(mR := Rotation_Matrix, dRoll => euler.A, dPitch => euler.B, dYaw => euler.C);

END_FUNCTION_BLOCK

// Device/Application/Topics_Vis
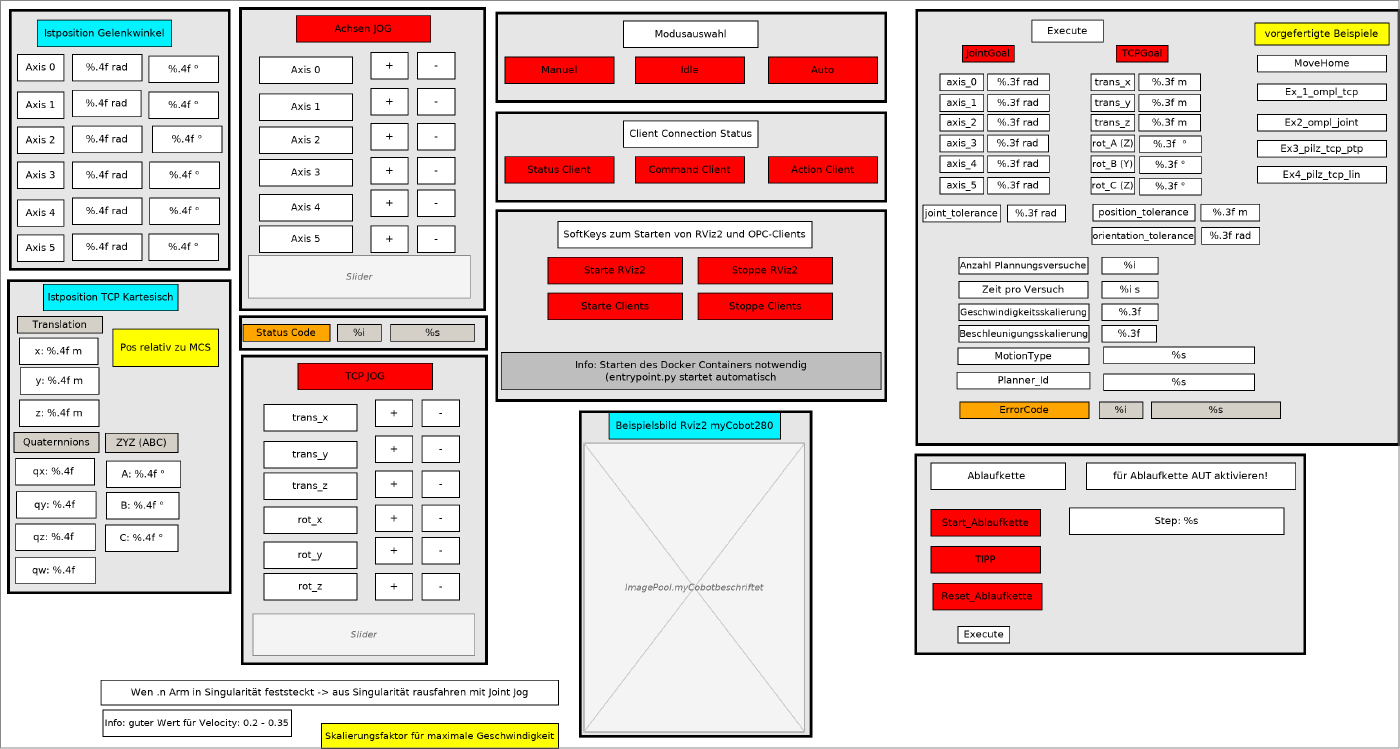
VISUALIZATION Topics_Vis  // 1557x834
    Rectangle (266,351 276x39)
    Rectangle (266,8 274x338)
    Rectangle (644,457 259x364)
    Rectangle (551,233 435x214)
    Rectangle (8,311 249x350)
    Rectangle (1018,10 539x486)
    Rectangle (551,13 435x101)
    Rectangle (10,10 246x291)
    Rectangle (41,22 150x30), "Istposition Gelenkwinkel"
    Rectangle (48,316 150x30), "Istposition TCP Kartesisch"
    Rectangle (21,376 88x30), "x: %.4f m", text variable: MAIN_PRG.RobotStatus.tcp_pose.trans_x
    Rectangle (22,409 88x30), "y: %.4f m", text variable: MAIN_PRG.RobotStatus.tcp_pose.trans_y
    Rectangle (21,445 89x30), "z: %.4f m", text variable: MAIN_PRG.RobotStatus.tcp_pose.trans_z
    Rectangle (17,510 88x30), "qx: %.4f", text variable: MAIN_PRG.RobotStatus.tcp_pose.rot_x
    Rectangle (18,547 89x30), "qy: %.4f", text variable: MAIN_PRG.RobotStatus.tcp_pose.rot_y
    Rectangle (17,583 89x30), "qz: %.4f", text variable: MAIN_PRG.RobotStatus.tcp_pose.rot_z
    Rectangle (17,620 89x30), "qw: %.4f", text variable: MAIN_PRG.RobotStatus.tcp_pose.rot_w
    Rectangle (412,58 42x30), "+"
        OnMouseDown: execute { MAIN_PRG.RobotCommand.axis_0 := +1; }
        OnMouseUp: execute { MAIN_PRG.RobotCommand.axis_0 := 0; }
    Rectangle (464,58 42x30), "-"
        OnMouseDown: execute { MAIN_PRG.RobotCommand.axis_0 := -1; }
        OnMouseUp: execute { MAIN_PRG.RobotCommand.axis_0 := 0; }
    Rectangle (412,98 42x30), "+"
        OnMouseDown: execute { MAIN_PRG.RobotCommand.axis_1 := +1; }
        OnMouseUp: execute { MAIN_PRG.RobotCommand.axis_1 := 0; }
    Rectangle (464,137 42x30), "-"
        OnMouseDown: execute { MAIN_PRG.RobotCommand.axis_2 := -1; }
        OnMouseUp: execute { MAIN_PRG.RobotCommand.axis_2 := 0; }
    Rectangle (412,137 42x30), "+"
        OnMouseDown: execute { MAIN_PRG.RobotCommand.axis_2 := +1; }
        OnMouseUp: execute { MAIN_PRG.RobotCommand.axis_2 := 0; }
    Rectangle (412,175 42x30), "+"
        OnMouseDown: execute { MAIN_PRG.RobotCommand.axis_3 := +1; }
        OnMouseUp: execute { MAIN_PRG.RobotCommand.axis_3 := 0; }
    Rectangle (464,98 42x30), "-"
        OnMouseDown: execute { MAIN_PRG.RobotCommand.axis_1 := -1; }
        OnMouseUp: execute { MAIN_PRG.RobotCommand.axis_1 := 0; }
    Rectangle (464,175 42x30), "-"
        OnMouseDown: execute { MAIN_PRG.RobotCommand.axis_3 := -1; }
        OnMouseUp: execute { MAIN_PRG.RobotCommand.axis_3 := 0; }
    Rectangle (412,211 42x30), "+"
        OnMouseDown: execute { MAIN_PRG.RobotCommand.axis_4 := +1; }
        OnMouseUp: execute { MAIN_PRG.RobotCommand.axis_4 := 0; }
    Rectangle (464,211 42x30), "-"
        OnMouseDown: execute { MAIN_PRG.RobotCommand.axis_4 := -1; }
        OnMouseUp: execute { MAIN_PRG.RobotCommand.axis_4 := 0; }
    Rectangle (412,251 42x30), "+"
        OnMouseDown: execute { MAIN_PRG.RobotCommand.axis_5 := +1; }
        OnMouseUp: execute { MAIN_PRG.RobotCommand.axis_5 := 0; }
    Rectangle (464,251 42x30), "-"
        OnMouseDown: execute { MAIN_PRG.RobotCommand.axis_5 := -1; }
        OnMouseUp: execute { MAIN_PRG.RobotCommand.axis_5 := 0; }
    Slider (276,284 247x48), variable: MAIN_PRG.RobotCommand.axis_velocity, scale 0..1
    Rectangle (693,23 150x30), "Modusauswahl"
    Rectangle (80,60 78x30), "%.4f rad", text variable: MAIN_PRG.RobotStatus.axis_pose.axis_0
    Rectangle (80,100 77x30), "%.4f rad", text variable: MAIN_PRG.RobotStatus.axis_pose.axis_1
    Rectangle (80,140 78x30), "%.4f rad", text variable: MAIN_PRG.RobotStatus.axis_pose.axis_2
    Rectangle (80,180 78x30), "%.4f rad", text variable: MAIN_PRG.RobotStatus.axis_pose.axis_3
    Rectangle (80,220 78x30), "%.4f rad", text variable: MAIN_PRG.RobotStatus.axis_pose.axis_4
    Rectangle (80,260 78x30), "%.4f rad", text variable: MAIN_PRG.RobotStatus.axis_pose.axis_5
    Rectangle (329,17 150x30), "Achsen JOG", colour toggle: GVL_OPCUA.RobotCommand.Mode_Axis
        toggle GVL_OPCUA.RobotCommand.Mode_Axis
        OnMouseClick: execute { GVL_OPCUA.RobotCommand.Mode_TCP := FALSE; }
    Rectangle (561,63 122x30), "Manuel", colour toggle: MAIN_PRG.Modes.MANUEL
        toggle MAIN_PRG.Modes.SEL_MAN p2164770859=TRUE
    Rectangle (854,63 122x30), "Auto", colour toggle: MAIN_PRG.Modes.AUTO
        toggle MAIN_PRG.Modes.SEL_AUTO p2164770859=TRUE
    Rectangle (706,63 122x30), "Idle", colour toggle: MAIN_PRG.Modes.IDLE
    Rectangle (1045,82 49x19), "axis_0"
    Rectangle (1045,105 49x19), "axis_1"
    Rectangle (1045,127 49x19), "axis_2"
    Rectangle (1045,150 49x19), "axis_3"
    Rectangle (1045,173 49x19), "axis_4"
    Rectangle (1045,197 49x19), "axis_5"
    Rectangle (1098,82 69x19), "%.3f rad", text variable: MAIN_PRG.RobotAction.axis_0
        OnMouseClick: write the text variable via Default
    Rectangle (1098,105 69x19), "%.3f rad", text variable: MAIN_PRG.RobotAction.axis_1
        OnMouseClick: write the text variable via Default
    Rectangle (1098,127 69x19), "%.3f rad", text variable: MAIN_PRG.RobotAction.axis_2
        OnMouseClick: write the text variable via Default
    Rectangle (1098,150 68x19), "%.3f rad", text variable: MAIN_PRG.RobotAction.axis_3
        OnMouseClick: write the text variable via Default
    Rectangle (1098,173 69x19), "%.3f rad", text variable: MAIN_PRG.RobotAction.axis_4
        OnMouseClick: write the text variable via Default
    Rectangle (1098,197 69x19), "%.3f rad", text variable: MAIN_PRG.RobotAction.axis_5
        OnMouseClick: write the text variable via Default
    Rectangle (1213,82 49x19), "trans_x"
    Rectangle (1213,105 49x19), "trans_y"
    Rectangle (1213,127 49x19), "trans_z"
    Rectangle (1266,82 69x19), "%.3f m", text variable: MAIN_PRG.RobotAction.trans_x
        OnMouseClick: write the text variable via Default
    Rectangle (1266,105 69x19), "%.3f m", text variable: MAIN_PRG.RobotAction.trans_y
        OnMouseClick: write the text variable via Default
    Rectangle (1266,127 69x19), "%.3f m", text variable: MAIN_PRG.RobotAction.trans_z
        OnMouseClick: write the text variable via Default
    Rectangle (1147,22 80x25), "Execute"
        tap GVL_OPCUA.Execute
    Rectangle (1070,50 58x19), "JointGoal", colour toggle: MAIN_PRG.RobotAction.Joint_Goal
        toggle MAIN_PRG.RobotAction.Joint_Goal
    Rectangle (1241,50 58x19), "TCPGoal", colour toggle: MAIN_PRG.RobotAction.TCP_Goal
        toggle MAIN_PRG.RobotAction.TCP_Goal
    Rectangle (1066,286 144x19), "Anzahl Plannungsversuche"
    Rectangle (1066,313 144x19), "Zeit pro Versuch"
    Rectangle (1066,338 145x19), "Geschwindigkeitsskalierung"
    Rectangle (1066,362 145x19), "Beschleunigungsskalierung"
    Rectangle (1215,227 114x19), "position_tolerance"
    Rectangle (1214,253 115x19), "orientation_tolerance"
    Rectangle (1225,286 63x19), "%i", text variable: MAIN_PRG.RobotAction.num_planning_attempts
        OnMouseClick: write the text variable via Default
    Rectangle (1225,313 63x19), "%i s", text variable: MAIN_PRG.RobotAction.allowed_planning_time
        OnMouseClick: write the text variable via Default
    Rectangle (1225,338 63x19), "%.3f", text variable: MAIN_PRG.RobotAction.max_velocity_scaling
        OnMouseClick: write the text variable via Default
    Rectangle (1225,362 61x19), "%.3f", text variable: MAIN_PRG.RobotAction.max_acceleration_scaling
        OnMouseClick: write the text variable via Default
    Rectangle (1335,227 66x19), "%.3f m", text variable: MAIN_PRG.RobotAction.position_tolerance
        OnMouseClick: write the text variable via Default
    Rectangle (1336,253 65x19), "%.3f rad", text variable: MAIN_PRG.RobotAction.orientation_tolerance
        OnMouseClick: write the text variable via Default
    Rectangle (1065,387 146x19), "MotionType"
    Rectangle (1064,414 148x19), "Planner_Id"
    Rectangle (1067,447 144x19), "ErrorCode"
    Rectangle (1222,447 49x19), "%i", text variable: MAIN_PRG.RobotAction.error_code
    Rectangle (1227,386 168x19), "%s", text variable: MAIN_PRG.RobotAction.Motion_Type
        OnMouseClick: write the text variable via Default
    Rectangle (1227,416 168x19), "%s", text variable: MAIN_PRG.RobotAction.Planner_ID
        OnMouseClick: write the text variable via Default
    Rectangle (1398,61 144x19), "MoveHome"
        tap MAIN_PRG.xMoveHome
    Rectangle (1280,447 144x19), "%s", text variable: MAIN_PRG.Status_Error_Codes_Action
    Rectangle (551,124 435x101)
    Rectangle (693,134 150x30), "Client Connection Status"
    Rectangle (561,174 122x30), "Status Client", colour toggle: MAIN_PRG.RobotStatus.client_connected
    Rectangle (854,174 122x30), "Action Client", colour toggle: MAIN_PRG.RobotAction.client_connected
    Rectangle (706,174 122x30), "Command Client", colour toggle: MAIN_PRG.RobotCommand.client_connected
    Rectangle (1398,93 144x19), "Ex_1_ompl_tcp"
        tap MAIN_PRG.xEx1_ompl_tcp
    Rectangle (1398,127 144x19), "Ex2_ompl_joint"
        tap MAIN_PRG.xEx2_ompl_joint
    Rectangle (1398,156 144x19), "Ex3_pilz_tcp_ptp"
        tap MAIN_PRG.xEx3_pilz_tcp_ptp
    Rectangle (1398,185 144x19), "Ex4_pilz_tcp_lin"
        tap MAIN_PRG.xEx4_pilz_tcp_lin
    Rectangle (165,62 78x30), "%.4f °", text variable: MAIN_PRG.RobotStatus.axis_pose.axis_0 *(180.0/GVL_OPCUA.PI)
    Rectangle (165,102 78x30), "%.4f °", text variable: MAIN_PRG.RobotStatus.axis_pose.axis_1 *(180.0/GVL_OPCUA.PI)
    Rectangle (169,140 78x30), "%.4f °", text variable: MAIN_PRG.RobotStatus.axis_pose.axis_2 *(180.0/GVL_OPCUA.PI)
    Rectangle (166,180 78x30), "%.4f °", text variable: MAIN_PRG.RobotStatus.axis_pose.axis_3 *(180.0/GVL_OPCUA.PI)
    Rectangle (166,220 78x30), "%.4f °", text variable: MAIN_PRG.RobotStatus.axis_pose.axis_4 *(180.0/GVL_OPCUA.PI)
    Rectangle (165,260 78x30), "%.4f °", text variable: MAIN_PRG.RobotStatus.axis_pose.axis_5 *(180.0/GVL_OPCUA.PI)
    Rectangle (118,513 83x30), "A: %.4f °", text variable: MAIN_PRG.Status_Quat_to_ZYZ.euler.A
    Rectangle (118,548 81x30), "B: %.4f °", text variable: MAIN_PRG.Status_Quat_to_ZYZ.euler.B
    Rectangle (117,584 81x30), "C: %.4f °", text variable: MAIN_PRG.Status_Quat_to_ZYZ.euler.C
    Rectangle (117,482 81x22), "ZYZ (ABC)"
    Rectangle (1017,505 435x224)
    Rectangle (1035,515 150x30), "Ablaufkette"
    Rectangle (1035,608 122x30), "TIPP", colour toggle: MAIN_PRG.RobotStatus.client_connected
        tap GVL_OPCUA.TIPP
    Rectangle (1035,567 122x30), "Start_Ablaufkette", colour toggle: MAIN_PRG.RobotStatus.client_connected
        tap GVL_OPCUA.Start_Ablaufkette
    Rectangle (1189,565 239x30), "Step: %s", text variable: Ablaufkette.SFCCurrentStep
    Rectangle (1208,515 233x30), "für Ablaufkette AUT aktivieren!"
    Rectangle (1037,649 122x30), "Reset_Ablaufkette", colour toggle: MAIN_PRG.RobotStatus.client_connected
        tap GVL_OPCUA.Reset_Ablaufkette
    Rectangle (1065,697 58x19), "Execute"
        tap GVL_OPCUA.Execute
    Rectangle (15,481 95x23), "Quaternnions"
    Rectangle (609,286 150x30), "Starte RViz2"
        toggle GVL_OPCUA.Start_RViz2
    Rectangle (609,326 150x30), "Starte Clients"
        toggle GVL_OPCUA.Start_OPCClients
    Rectangle (776,326 150x30), "Stoppe Clients"
        toggle GVL_OPCUA.Stop_OPC_Clients
    Rectangle (776,286 150x30), "Stoppe RViz2"
        toggle GVL_OPCUA.Stop_RViz2
    Rectangle (288,63 104x30), "Axis 0"
    Rectangle (288,104 104x30), "Axis 1"
    Rectangle (288,141 104x30), "Axis 2"
    Rectangle (288,177 104x30), "Axis 3"
    Rectangle (288,216 104x30), "Axis 4"
    Rectangle (288,251 104x30), "Axis 5"
    Rectangle (19,60 52x30), "Axis 0"
    Rectangle (19,102 52x30), "Axis 1"
    Rectangle (19,141 52x30), "Axis 2"
    Rectangle (19,180 52x30), "Axis 3"
    Rectangle (19,222 52x30), "Axis 4"
    Rectangle (19,261 52x30), "Axis 5"
    RoundedRectangle (125,366 118x42), "Pos relativ zu MCS"
    Image (649,493 246x322), image: ImagePool.myCobotbeschriftet
    Rectangle (677,459 191x30), "Beispielsbild Rviz2 myCobot280"
    RoundedRectangle (1395,25 150x25), "vorgefertigte Beispiele"
    Rectangle (620,246 283x30), "SoftKeys zum Starten von RViz2 und OPC-Clients"
    Rectangle (557,392 423x42), "Info: Starten des Docker Containers notwendig (entrypoint.py startet automatisch"
    Rectangle (1213,150 49x19), "rot_A (Z)"
    Rectangle (1213,173 49x19), "rot_B (Y)"
    Rectangle (1213,197 49x19), "rot_C (Z)"
    Rectangle (1267,151 69x19), "%.3f °", text variable: GVL_OPCUA.rot_A
        OnMouseClick: write the text variable via Default
    Rectangle (1267,174 69x19), "%.3f °", text variable: GVL_OPCUA.rot_B
        OnMouseClick: write the text variable via Default
    Rectangle (1267,198 69x19), "%.3f °", text variable: GVL_OPCUA.rot_C
        OnMouseClick: write the text variable via Default
    Rectangle (1026,228 87x19), "joint_tolerance"
    Rectangle (1120,228 65x19), "%.3f rad", text variable: MAIN_PRG.RobotAction.joint_tolerance
        OnMouseClick: write the text variable via Default
    Rectangle (268,395 274x345)
    Rectangle (417,445 42x30), "+"
        OnMouseDown: execute { MAIN_PRG.RobotCommand.trans_x := +1; }
        OnMouseUp: execute { MAIN_PRG.RobotCommand.trans_x := 0; }
    Rectangle (469,445 42x30), "-"
        OnMouseDown: execute { MAIN_PRG.RobotCommand.trans_x := -1; }
        OnMouseUp: execute { MAIN_PRG.RobotCommand.trans_x := 0; }
    Rectangle (417,485 42x30), "+"
        OnMouseDown: execute { MAIN_PRG.RobotCommand.trans_y := +1; }
        OnMouseUp: execute { MAIN_PRG.RobotCommand.trans_y := 0; }
    Rectangle (469,524 42x30), "-"
        OnMouseDown: execute { MAIN_PRG.RobotCommand.trans_z := -1; }
        OnMouseUp: execute { MAIN_PRG.RobotCommand.trans_z := 0; }
    Rectangle (417,524 42x30), "+"
        OnMouseDown: execute { MAIN_PRG.RobotCommand.trans_z := +1; }
        OnMouseUp: execute { MAIN_PRG.RobotCommand.trans_z := 0; }
    Rectangle (417,562 42x30), "+"
        OnMouseDown: execute { MAIN_PRG.RobotCommand.rot_x := +1; }
        OnMouseUp: execute { MAIN_PRG.RobotCommand.rot_x := 0; }
    Rectangle (469,485 42x30), "-"
        OnMouseDown: execute { MAIN_PRG.RobotCommand.trans_y := -1; }
        OnMouseUp: execute { MAIN_PRG.RobotCommand.trans_y := 0; }
    Rectangle (469,562 42x30), "-"
        OnMouseDown: execute { MAIN_PRG.RobotCommand.rot_x := -1; }
        OnMouseUp: execute { MAIN_PRG.RobotCommand.rot_x := 0; }
    Rectangle (417,598 42x30), "+"
        OnMouseDown: execute { MAIN_PRG.RobotCommand.rot_y := +1; }
        OnMouseUp: execute { MAIN_PRG.RobotCommand.rot_y := 0; }
    Rectangle (469,598 42x30), "-"
        OnMouseDown: execute { MAIN_PRG.RobotCommand.rot_y := -1; }
        OnMouseUp: execute { MAIN_PRG.RobotCommand.rot_y := 0; }
    Rectangle (417,638 42x30), "+"
        OnMouseDown: execute { MAIN_PRG.RobotCommand.rot_z := +1; }
        OnMouseUp: execute { MAIN_PRG.RobotCommand.rot_z := 0; }
    Rectangle (469,638 42x30), "-"
        OnMouseDown: execute { MAIN_PRG.RobotCommand.rot_z := -1; }
        OnMouseUp: execute { MAIN_PRG.RobotCommand.rot_z := 0; }
    Slider (281,683 247x47), variable: MAIN_PRG.RobotCommand.tcp_velocity, scale 0..1
    Rectangle (331,404 150x30), "TCP JOG", colour toggle: GVL_OPCUA.RobotCommand.Mode_TCP
        toggle GVL_OPCUA.RobotCommand.Mode_TCP
        OnMouseClick: execute { GVL_OPCUA.RobotCommand.Mode_Axis := FALSE; }
    Rectangle (293,450 104x30), "trans_x"
    Rectangle (293,491 104x30), "trans_y"
    Rectangle (293,526 104x30), "trans_z"
    Rectangle (293,564 104x30), "rot_x"
    Rectangle (293,603 104x30), "rot_y"
    Rectangle (293,638 104x30), "rot_z"
    Rectangle (114,790 210x30), "Info: guter Wert für Velocity: 0.2 - 0.35"
    Rectangle (112,757 509x28), "Wen .n Arm in Singularität feststeckt -> aus Singularität rausfahren mit Joint Jog"
    Rectangle (270,361 97x19), "Status Code"
    Rectangle (375,361 49x19), "%i", text variable: MAIN_PRG.RobotCommand.status
    Rectangle (434,361 94x19), "%s", text variable: MAIN_PRG.Status_Servo
    Rectangle (19,352 95x19), "Translation"
    RoundedRectangle (357,805 264x29), "Skalierungsfaktor für maximale Geschwindigkeit"
END_VISUALIZATION

// Device/Application/VISU_Auto
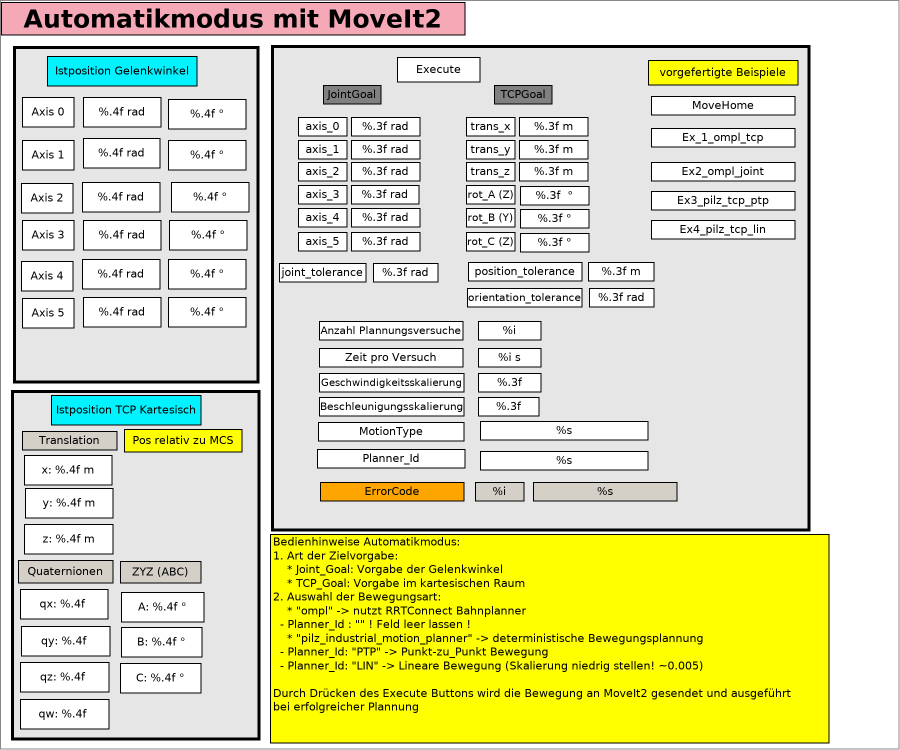
VISUALIZATION VISU_Auto  // 900x750
    Rectangle (271,45 539x486)
    Rectangle (298,117 49x19), "axis_0"
    Rectangle (298,140 49x19), "axis_1"
    Rectangle (298,162 49x19), "axis_2"
    Rectangle (298,185 49x19), "axis_3"
    Rectangle (298,208 49x19), "axis_4"
    Rectangle (298,232 49x19), "axis_5"
    Rectangle (351,117 69x19), "%.3f rad", text variable: GVL_OPCUA.axis_0
        OnMouseClick: write the text variable via Default
    Rectangle (351,140 69x19), "%.3f rad", text variable: GVL_OPCUA.axis_1
        OnMouseClick: write the text variable via Default
    Rectangle (351,162 69x19), "%.3f rad", text variable: GVL_OPCUA.axis_2
        OnMouseClick: write the text variable via Default
    Rectangle (351,185 68x19), "%.3f rad", text variable: GVL_OPCUA.axis_3
        OnMouseClick: write the text variable via Default
    Rectangle (351,208 69x19), "%.3f rad", text variable: GVL_OPCUA.axis_4
        OnMouseClick: write the text variable via Default
    Rectangle (351,232 69x19), "%.3f rad", text variable: GVL_OPCUA.axis_5
        OnMouseClick: write the text variable via Default
    Rectangle (466,117 49x19), "trans_x"
    Rectangle (466,140 49x19), "trans_y"
    Rectangle (466,162 49x19), "trans_z"
    Rectangle (519,117 69x19), "%.3f m", text variable: GVL_OPCUA.trans_x
        OnMouseClick: write the text variable via Default
    Rectangle (519,140 69x19), "%.3f m", text variable: GVL_OPCUA.trans_y
        OnMouseClick: write the text variable via Default
    Rectangle (519,162 69x19), "%.3f m", text variable: GVL_OPCUA.trans_z
        OnMouseClick: write the text variable via Default
    Rectangle (397,57 83x25), "Execute"
        tap GVL_OPCUA.Execute
    Rectangle (323,85 58x19), "JointGoal", colour toggle: GVL_OPCUA.Joint_Goal
        toggle GVL_OPCUA.Joint_Goal
    Rectangle (494,85 58x19), "TCPGoal", colour toggle: GVL_OPCUA.TCP_GOAL
        toggle GVL_OPCUA.TCP_GOAL
    Rectangle (319,321 144x19), "Anzahl Plannungsversuche"
    Rectangle (319,348 144x19), "Zeit pro Versuch"
    Rectangle (319,373 145x19), "Geschwindigkeitsskalierung"
    Rectangle (319,397 145x19), "Beschleunigungsskalierung"
    Rectangle (468,262 114x19), "position_tolerance"
    Rectangle (467,288 115x19), "orientation_tolerance"
    Rectangle (478,321 63x19), "%i", text variable: GVL_OPCUA.num_planning_attempts
        OnMouseClick: write the text variable via Default
    Rectangle (478,348 63x19), "%i s", text variable: GVL_OPCUA.allowed_planning_time
        OnMouseClick: write the text variable via Default
    Rectangle (478,373 63x19), "%.3f", text variable: GVL_OPCUA.max_velocity_scaling
        OnMouseClick: write the text variable via Default
    Rectangle (478,397 61x19), "%.3f", text variable: GVL_OPCUA.max_acceleration_scaling
        OnMouseClick: write the text variable via Default
    Rectangle (588,262 66x19), "%.3f m", text variable: GVL_OPCUA.position_tolerance
        OnMouseClick: write the text variable via Default
    Rectangle (589,288 65x19), "%.3f rad", text variable: GVL_OPCUA.orientation_tolerance
        OnMouseClick: write the text variable via Default
    Rectangle (318,422 146x19), "MotionType"
    Rectangle (317,449 148x19), "Planner_Id"
    Rectangle (320,482 144x19), "ErrorCode"
    Rectangle (475,482 49x19), "%i", text variable: MAIN_PRG.RobotAction.error_code
    Rectangle (480,421 168x19), "%s", text variable: GVL_OPCUA.Motion_Type
        OnMouseClick: write the text variable via Default
    Rectangle (480,451 168x19), "%s", text variable: GVL_OPCUA.Planner_ID
        OnMouseClick: write the text variable via Default
    Rectangle (651,96 144x19), "MoveHome"
        tap MAIN_PRG.xMoveHome
    Rectangle (533,482 144x19), "%s", text variable: MAIN_PRG.Status_Error_Codes_Action
    Rectangle (651,128 144x19), "Ex_1_ompl_tcp"
        tap MAIN_PRG.xEx1_ompl_tcp
    Rectangle (651,162 144x19), "Ex2_ompl_joint"
        tap MAIN_PRG.xEx2_ompl_joint
    Rectangle (651,191 144x19), "Ex3_pilz_tcp_ptp"
        tap MAIN_PRG.xEx3_pilz_tcp_ptp
    Rectangle (651,220 144x19), "Ex4_pilz_tcp_lin"
        tap MAIN_PRG.xEx4_pilz_tcp_lin
    RoundedRectangle (648,60 150x25), "vorgefertigte Beispiele"
    Rectangle (466,185 49x19), "rot_A (Z)"
    Rectangle (466,208 49x19), "rot_B (Y)"
    Rectangle (466,232 49x19), "rot_C (Z)"
    Rectangle (520,186 69x19), "%.3f °", text variable: GVL_OPCUA.rot_A
        OnMouseClick: write the text variable via Default
    Rectangle (520,209 69x19), "%.3f °", text variable: GVL_OPCUA.rot_B
        OnMouseClick: write the text variable via Default
    Rectangle (520,233 69x19), "%.3f °", text variable: GVL_OPCUA.rot_C
        OnMouseClick: write the text variable via Default
    Rectangle (279,263 87x19), "joint_tolerance"
    Rectangle (373,263 65x19), "%.3f rad", text variable: GVL_OPCUA.joint_tolerance
        OnMouseClick: write the text variable via Default
    Rectangle (11,390 249x350)
    Rectangle (13,46 246x337)
    Rectangle (47,56 150x30), "Istposition Gelenkwinkel"
    Rectangle (51,395 150x30), "Istposition TCP Kartesisch"
    Rectangle (24,455 88x30), "x: %.4f m", text variable: GVL_OPCUA.RobotStatus.Ist_Pos_TCP.trans_x
    Rectangle (25,488 88x30), "y: %.4f m", text variable: GVL_OPCUA.RobotStatus.Ist_Pos_TCP.trans_y
    Rectangle (24,524 89x30), "z: %.4f m", text variable: GVL_OPCUA.RobotStatus.Ist_Pos_TCP.trans_z
    Rectangle (20,589 88x30), "qx: %.4f", text variable: GVL_OPCUA.RobotStatus.Ist_Pos_TCP.rot_x
    Rectangle (21,626 89x30), "qy: %.4f", text variable: GVL_OPCUA.RobotStatus.Ist_Pos_TCP.rot_y
    Rectangle (20,662 89x30), "qz: %.4f", text variable: GVL_OPCUA.RobotStatus.Ist_Pos_TCP.rot_z
    Rectangle (20,699 89x30), "qw: %.4f", text variable: GVL_OPCUA.RobotStatus.Ist_Pos_TCP.rot_w
    Rectangle (83,97 78x30), "%.4f rad", text variable: GVL_OPCUA.RobotStatus.Ist_Pos_Axis.axis_0
    Rectangle (83,138 77x30), "%.4f rad", text variable: GVL_OPCUA.RobotStatus.Ist_Pos_Axis.axis_1
    Rectangle (82,182 78x30), "%.4f rad", text variable: GVL_OPCUA.RobotStatus.Ist_Pos_Axis.axis_2
    Rectangle (83,220 78x30), "%.4f rad", text variable: GVL_OPCUA.RobotStatus.Ist_Pos_Axis.axis_3
    Rectangle (82,259 78x30), "%.4f rad", text variable: GVL_OPCUA.RobotStatus.Ist_Pos_Axis.axis_4
    Rectangle (83,297 78x30), "%.4f rad", text variable: GVL_OPCUA.RobotStatus.Ist_Pos_Axis.axis_5
    Rectangle (168,99 78x30), "%.4f °", text variable: GVL_OPCUA.RobotStatus.Ist_Pos_Axis.axis_0 *(180.0/GVL_OPCUA.PI)
    Rectangle (168,140 78x30), "%.4f °", text variable: GVL_OPCUA.RobotStatus.Ist_Pos_Axis.axis_1 *(180.0/GVL_OPCUA.PI)
    Rectangle (171,182 78x30), "%.4f °", text variable: GVL_OPCUA.RobotStatus.Ist_Pos_Axis.axis_2 *(180.0/GVL_OPCUA.PI)
    Rectangle (169,220 78x30), "%.4f °", text variable: GVL_OPCUA.RobotStatus.Ist_Pos_Axis.axis_3 *(180.0/GVL_OPCUA.PI)
    Rectangle (168,259 78x30), "%.4f °", text variable: GVL_OPCUA.RobotStatus.Ist_Pos_Axis.axis_4 *(180.0/GVL_OPCUA.PI)
    Rectangle (168,297 78x30), "%.4f °", text variable: GVL_OPCUA.RobotStatus.Ist_Pos_Axis.axis_5 *(180.0/GVL_OPCUA.PI)
    Rectangle (121,592 83x30), "A: %.4f °", text variable: MAIN_PRG.Status_Quat_to_ZYZ.euler.A
    Rectangle (121,627 81x30), "B: %.4f °", text variable: MAIN_PRG.Status_Quat_to_ZYZ.euler.B
    Rectangle (120,663 81x30), "C: %.4f °", text variable: MAIN_PRG.Status_Quat_to_ZYZ.euler.C
    Rectangle (120,561 81x22), "ZYZ (ABC)"
    Rectangle (18,560 95x23), "Quaternionen"
    Rectangle (22,97 52x30), "Axis 0"
    Rectangle (22,140 52x30), "Axis 1"
    Rectangle (21,183 52x30), "Axis 2"
    Rectangle (22,220 52x30), "Axis 3"
    Rectangle (21,261 52x30), "Axis 4"
    Rectangle (22,298 52x30), "Axis 5"
    RoundedRectangle (124,429 118x23), "Pos relativ zu MCS"
    Rectangle (22,431 95x19), "Translation"
    Rectangle (1,2 464x33), "Automatikmodus mit MoveIt2"
    RoundedRectangle (270,534 559x209), "Bedienhinweise Automatikmodus: 1. Art der Zielvorgabe: * Joint_Goal: Vorgabe der Gelenkwinkel * TCP_Goal: Vorgabe im kartesischen Raum 2. Auswahl der Bewegungsart: * "ompl" -> nutzt RRTConnect Bahnplanner - Planner_Id : "" ! Feld leer lassen ! * "pilz_industrial_motion_planner" -> deterministische Bewegungsplannung - Planner_Id: "PTP" -> Punkt-zu_Punkt Bewegung - Planner_Id: "LIN" -> Lineare Bewegung (Skalierung niedrig stellen! ~0.005) Durch Drücken des Execute Buttons wird die Bewegung an MoveIt2 gesendet und ausgeführt bei erfolgreicher Plannung"
END_VISUALIZATION

// Device/Application/VISU_Startseite
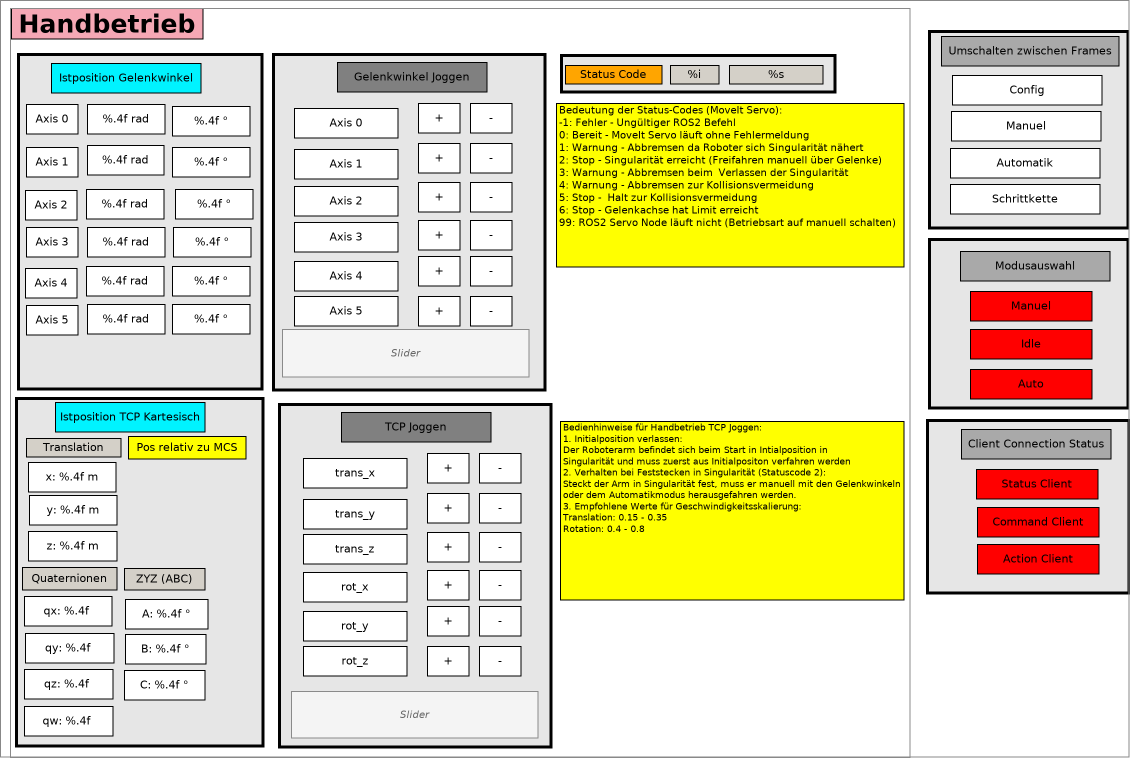
VISUALIZATION VISU_Startseite  // 1130x758
    Rectangle (928,30 201x199)
    Frame (10,8 900x750)
        shows VISU_Manuell()
        shows VISU_Konfig()
        shows VISU_Auto()
        shows VISU_Schrittkette()
    Rectangle (952,75 150x30), "Config"
        OnMouseClick: FrameSelectionChange Selection=SelectedFrame=848abb15-4fea-4ce4-a60a-73a186e6a183, Selection=1, GlobSel=AssignType=Directly, SelType=Locally, SelectionStep=SelectedAction=SwitchNext
    Rectangle (951,111 150x30), "Manuel"
        OnMouseClick: FrameSelectionChange Selection=SelectedFrame=848abb15-4fea-4ce4-a60a-73a186e6a183, GlobSel=AssignType=Directly, SelType=Locally, SelectionStep=SelectedAction=SwitchNext
    Rectangle (950,148 150x30), "Automatik"
        OnMouseClick: FrameSelectionChange Selection=SelectedFrame=848abb15-4fea-4ce4-a60a-73a186e6a183, Selection=2, GlobSel=AssignType=Directly, SelType=Locally, SelectionStep=SelectedAction=SwitchNext
    Rectangle (941,36 178x30), "Umschalten zwischen Frames"
    Rectangle (928,238 201x171)
    Rectangle (960,251 150x30), "Modusauswahl"
    Rectangle (970,291 122x30), "Manuel", colour toggle: MAIN_PRG.Modes.MANUEL
        toggle MAIN_PRG.Modes.SEL_MAN p2164770859=TRUE
    Rectangle (970,369 122x30), "Auto", colour toggle: MAIN_PRG.Modes.AUTO
        toggle MAIN_PRG.Modes.SEL_AUTO p2164770859=TRUE
    Rectangle (970,329 122x30), "Idle", colour toggle: MAIN_PRG.Modes.IDLE
    Rectangle (926,419 204x175)
    Rectangle (961,429 150x30), "Client Connection Status"
    Rectangle (976,469 122x30), "Status Client", colour toggle: MAIN_PRG.RobotStatus.client_connected
    Rectangle (977,544 122x30), "Action Client", colour toggle: MAIN_PRG.RobotAction.client_connected
    Rectangle (977,507 122x30), "Command Client", colour toggle: MAIN_PRG.RobotCommand.client_connected
    Rectangle (950,184 150x30), "Schrittkette"
        OnMouseClick: FrameSelectionChange Selection=SelectedFrame=848abb15-4fea-4ce4-a60a-73a186e6a183, Selection=3, GlobSel=AssignType=Directly, SelType=Locally, SelectionStep=SelectedAction=SwitchNext
END_VISUALIZATION

// Device/Application/VISU_Manuell
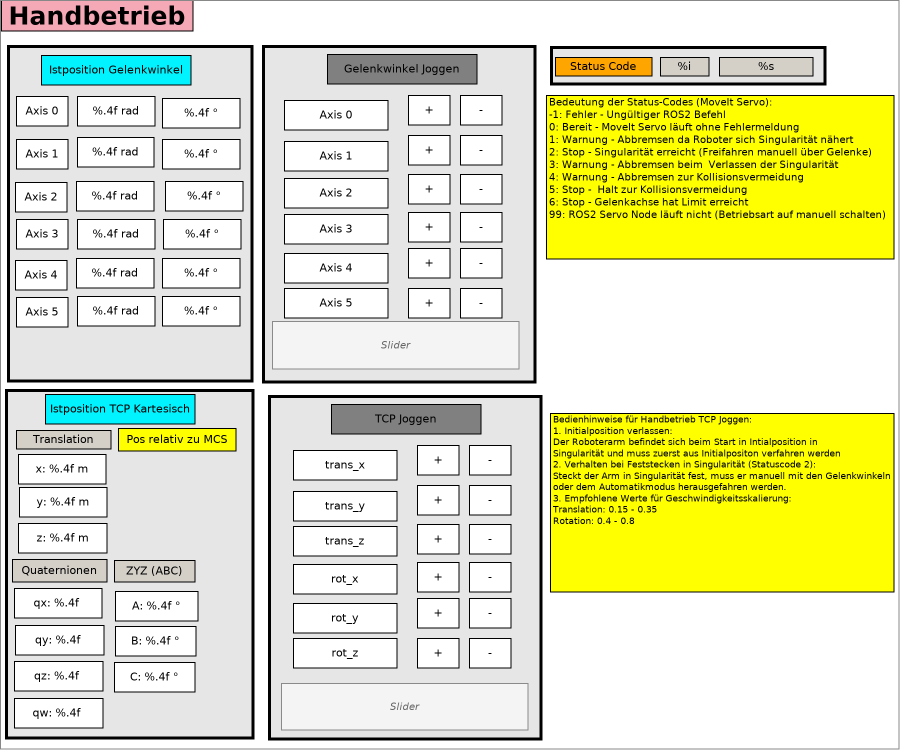
VISUALIZATION VISU_Manuell  // 900x750
    Rectangle (550,46 276x39)
    Rectangle (262,45 274x338)
    Rectangle (408,95 42x30), "+"
        OnMouseDown: execute { MAIN_PRG.RobotCommand.axis_0 := +1; }
        OnMouseUp: execute { MAIN_PRG.RobotCommand.axis_0 := 0; }
    Rectangle (460,95 42x30), "-"
        OnMouseDown: execute { MAIN_PRG.RobotCommand.axis_0 := -1; }
        OnMouseUp: execute { MAIN_PRG.RobotCommand.axis_0 := 0; }
    Rectangle (408,135 42x30), "+"
        OnMouseDown: execute { MAIN_PRG.RobotCommand.axis_1 := +1; }
        OnMouseUp: execute { MAIN_PRG.RobotCommand.axis_1 := 0; }
    Rectangle (460,174 42x30), "-"
        OnMouseDown: execute { MAIN_PRG.RobotCommand.axis_2 := -1; }
        OnMouseUp: execute { MAIN_PRG.RobotCommand.axis_2 := 0; }
    Rectangle (408,174 42x30), "+"
        OnMouseDown: execute { MAIN_PRG.RobotCommand.axis_2 := +1; }
        OnMouseUp: execute { MAIN_PRG.RobotCommand.axis_2 := 0; }
    Rectangle (408,212 42x30), "+"
        OnMouseDown: execute { MAIN_PRG.RobotCommand.axis_3 := +1; }
        OnMouseUp: execute { MAIN_PRG.RobotCommand.axis_3 := 0; }
    Rectangle (460,135 42x30), "-"
        OnMouseDown: execute { MAIN_PRG.RobotCommand.axis_1 := -1; }
        OnMouseUp: execute { MAIN_PRG.RobotCommand.axis_1 := 0; }
    Rectangle (460,212 42x30), "-"
        OnMouseDown: execute { MAIN_PRG.RobotCommand.axis_3 := -1; }
        OnMouseUp: execute { MAIN_PRG.RobotCommand.axis_3 := 0; }
    Rectangle (408,248 42x30), "+"
        OnMouseDown: execute { MAIN_PRG.RobotCommand.axis_4 := +1; }
        OnMouseUp: execute { MAIN_PRG.RobotCommand.axis_4 := 0; }
    Rectangle (460,248 42x30), "-"
        OnMouseDown: execute { MAIN_PRG.RobotCommand.axis_4 := -1; }
        OnMouseUp: execute { MAIN_PRG.RobotCommand.axis_4 := 0; }
    Rectangle (408,288 42x30), "+"
        OnMouseDown: execute { MAIN_PRG.RobotCommand.axis_5 := +1; }
        OnMouseUp: execute { MAIN_PRG.RobotCommand.axis_5 := 0; }
    Rectangle (460,288 42x30), "-"
        OnMouseDown: execute { MAIN_PRG.RobotCommand.axis_5 := -1; }
        OnMouseUp: execute { MAIN_PRG.RobotCommand.axis_5 := 0; }
    Slider (272,321 247x48), variable: MAIN_PRG.RobotCommand.axis_velocity, scale 0..1
    Rectangle (327,54 150x30), "Gelenkwinkel Joggen", colour toggle: GVL_OPCUA.RobotCommand.Mode_Axis
        toggle GVL_OPCUA.RobotCommand.Mode_Axis
        OnMouseClick: execute { GVL_OPCUA.RobotCommand.Mode_TCP := FALSE; }
    Rectangle (284,100 104x30), "Axis 0"
    Rectangle (284,141 104x30), "Axis 1"
    Rectangle (284,178 104x30), "Axis 2"
    Rectangle (284,214 104x30), "Axis 3"
    Rectangle (284,253 104x30), "Axis 4"
    Rectangle (284,288 104x30), "Axis 5"
    Rectangle (268,395 274x345)
    Rectangle (417,445 42x30), "+"
        OnMouseDown: execute { MAIN_PRG.RobotCommand.trans_x := +1; }
        OnMouseUp: execute { MAIN_PRG.RobotCommand.trans_x := 0; }
    Rectangle (469,445 42x30), "-"
        OnMouseDown: execute { MAIN_PRG.RobotCommand.trans_x := -1; }
        OnMouseUp: execute { MAIN_PRG.RobotCommand.trans_x := 0; }
    Rectangle (417,485 42x30), "+"
        OnMouseDown: execute { MAIN_PRG.RobotCommand.trans_y := +1; }
        OnMouseUp: execute { MAIN_PRG.RobotCommand.trans_y := 0; }
    Rectangle (469,524 42x30), "-"
        OnMouseDown: execute { MAIN_PRG.RobotCommand.trans_z := -1; }
        OnMouseUp: execute { MAIN_PRG.RobotCommand.trans_z := 0; }
    Rectangle (417,524 42x30), "+"
        OnMouseDown: execute { MAIN_PRG.RobotCommand.trans_z := +1; }
        OnMouseUp: execute { MAIN_PRG.RobotCommand.trans_z := 0; }
    Rectangle (417,562 42x30), "+"
        OnMouseDown: execute { MAIN_PRG.RobotCommand.rot_x := +1; }
        OnMouseUp: execute { MAIN_PRG.RobotCommand.rot_x := 0; }
    Rectangle (469,485 42x30), "-"
        OnMouseDown: execute { MAIN_PRG.RobotCommand.trans_y := -1; }
        OnMouseUp: execute { MAIN_PRG.RobotCommand.trans_y := 0; }
    Rectangle (469,562 42x30), "-"
        OnMouseDown: execute { MAIN_PRG.RobotCommand.rot_x := -1; }
        OnMouseUp: execute { MAIN_PRG.RobotCommand.rot_x := 0; }
    Rectangle (417,598 42x30), "+"
        OnMouseDown: execute { MAIN_PRG.RobotCommand.rot_y := +1; }
        OnMouseUp: execute { MAIN_PRG.RobotCommand.rot_y := 0; }
    Rectangle (469,598 42x30), "-"
        OnMouseDown: execute { MAIN_PRG.RobotCommand.rot_y := -1; }
        OnMouseUp: execute { MAIN_PRG.RobotCommand.rot_y := 0; }
    Rectangle (417,638 42x30), "+"
        OnMouseDown: execute { MAIN_PRG.RobotCommand.rot_z := +1; }
        OnMouseUp: execute { MAIN_PRG.RobotCommand.rot_z := 0; }
    Rectangle (469,638 42x30), "-"
        OnMouseDown: execute { MAIN_PRG.RobotCommand.rot_z := -1; }
        OnMouseUp: execute { MAIN_PRG.RobotCommand.rot_z := 0; }
    Slider (281,683 247x47), variable: MAIN_PRG.RobotCommand.tcp_velocity, scale 0..1
    Rectangle (331,404 150x30), "TCP Joggen", colour toggle: GVL_OPCUA.RobotCommand.Mode_TCP
        toggle GVL_OPCUA.RobotCommand.Mode_TCP
        OnMouseClick: execute { GVL_OPCUA.RobotCommand.Mode_Axis := FALSE; }
    Rectangle (293,450 104x30), "trans_x"
    Rectangle (293,491 104x30), "trans_y"
    Rectangle (293,526 104x30), "trans_z"
    Rectangle (293,564 104x30), "rot_x"
    Rectangle (293,603 104x30), "rot_y"
    Rectangle (293,638 104x30), "rot_z"
    Rectangle (555,57 97x19), "Status Code"
    Rectangle (660,57 49x19), "%i", text variable: MAIN_PRG.RobotCommand.status
    Rectangle (719,57 94x19), "%s", text variable: MAIN_PRG.Status_Servo
    Rectangle (1,0 192x31), "Handbetrieb"
    RoundedRectangle (550,413 344x179), "Bedienhinweise für Handbetrieb TCP Joggen: 1. Initialposition verlassen: Der Roboterarm befindet sich beim Start in Intialposition in Singularität und muss zuerst aus Initialpositon verfahren werden 2. Verhalten bei Feststecken in Singularität (Statuscode 2): Steckt der Arm in Singularität fest, muss er manuell mit den Gelenkwinkeln oder dem Automatikmodus herausgefahren werden. 3. Empfohlene Werte für Geschwindigkeitsskalierung: Translation: 0.15 - 0.35 Rotation: 0.4 - 0.8"
    RoundedRectangle (546,95 348x164), "Bedeutung der Status-Codes (MoveIt Servo): -1: Fehler - Ungültiger ROS2 Befehl 0: Bereit - MoveIt Servo läuft ohne Fehlermeldung 1: Warnung - Abbremsen da Roboter sich Singularität nähert 2: Stop - Singularität erreicht (Freifahren manuell über Gelenke) 3: Warnung - Abbremsen beim Verlassen der Singularität 4: Warnung - Abbremsen zur Kollisionsvermeidung 5: Stop - Halt zur Kollisionsvermeidung 6: Stop - Gelenkachse hat Limit erreicht 99: ROS2 Servo Node läuft nicht (Betriebsart auf manuell schalten)"
    Rectangle (5,389 249x350)
    Rectangle (7,45 246x337)
    Rectangle (41,55 150x30), "Istposition Gelenkwinkel"
    Rectangle (45,394 150x30), "Istposition TCP Kartesisch"
    Rectangle (18,454 88x30), "x: %.4f m", text variable: GVL_OPCUA.RobotStatus.Ist_Pos_TCP.trans_x
    Rectangle (19,487 88x30), "y: %.4f m", text variable: GVL_OPCUA.RobotStatus.Ist_Pos_TCP.trans_y
    Rectangle (18,523 89x30), "z: %.4f m", text variable: GVL_OPCUA.RobotStatus.Ist_Pos_TCP.trans_z
    Rectangle (14,588 88x30), "qx: %.4f", text variable: GVL_OPCUA.RobotStatus.Ist_Pos_TCP.rot_x
    Rectangle (15,625 89x30), "qy: %.4f", text variable: GVL_OPCUA.RobotStatus.Ist_Pos_TCP.rot_y
    Rectangle (14,661 89x30), "qz: %.4f", text variable: GVL_OPCUA.RobotStatus.Ist_Pos_TCP.rot_z
    Rectangle (14,698 89x30), "qw: %.4f", text variable: GVL_OPCUA.RobotStatus.Ist_Pos_TCP.rot_w
    Rectangle (77,96 78x30), "%.4f rad", text variable: GVL_OPCUA.RobotStatus.Ist_Pos_Axis.axis_0
    Rectangle (77,137 77x30), "%.4f rad", text variable: GVL_OPCUA.RobotStatus.Ist_Pos_Axis.axis_1
    Rectangle (76,181 78x30), "%.4f rad", text variable: GVL_OPCUA.RobotStatus.Ist_Pos_Axis.axis_2
    Rectangle (77,219 78x30), "%.4f rad", text variable: GVL_OPCUA.RobotStatus.Ist_Pos_Axis.axis_3
    Rectangle (76,258 78x30), "%.4f rad", text variable: GVL_OPCUA.RobotStatus.Ist_Pos_Axis.axis_4
    Rectangle (77,296 78x30), "%.4f rad", text variable: GVL_OPCUA.RobotStatus.Ist_Pos_Axis.axis_5
    Rectangle (162,98 78x30), "%.4f °", text variable: GVL_OPCUA.RobotStatus.Ist_Pos_Axis.axis_0 *(180.0/GVL_OPCUA.PI)
    Rectangle (162,139 78x30), "%.4f °", text variable: GVL_OPCUA.RobotStatus.Ist_Pos_Axis.axis_1 *(180.0/GVL_OPCUA.PI)
    Rectangle (165,181 78x30), "%.4f °", text variable: GVL_OPCUA.RobotStatus.Ist_Pos_Axis.axis_2 *(180.0/GVL_OPCUA.PI)
    Rectangle (163,219 78x30), "%.4f °", text variable: GVL_OPCUA.RobotStatus.Ist_Pos_Axis.axis_3 *(180.0/GVL_OPCUA.PI)
    Rectangle (162,258 78x30), "%.4f °", text variable: GVL_OPCUA.RobotStatus.Ist_Pos_Axis.axis_4 *(180.0/GVL_OPCUA.PI)
    Rectangle (162,296 78x30), "%.4f °", text variable: GVL_OPCUA.RobotStatus.Ist_Pos_Axis.axis_5 *(180.0/GVL_OPCUA.PI)
    Rectangle (115,591 83x30), "A: %.4f °", text variable: MAIN_PRG.Status_Quat_to_ZYZ.euler.A
    Rectangle (115,626 81x30), "B: %.4f °", text variable: MAIN_PRG.Status_Quat_to_ZYZ.euler.B
    Rectangle (114,662 81x30), "C: %.4f °", text variable: MAIN_PRG.Status_Quat_to_ZYZ.euler.C
    Rectangle (114,560 81x22), "ZYZ (ABC)"
    Rectangle (12,559 95x23), "Quaternionen"
    Rectangle (16,96 52x30), "Axis 0"
    Rectangle (16,139 52x30), "Axis 1"
    Rectangle (15,182 52x30), "Axis 2"
    Rectangle (16,219 52x30), "Axis 3"
    Rectangle (15,260 52x30), "Axis 4"
    Rectangle (16,297 52x30), "Axis 5"
    RoundedRectangle (118,428 118x23), "Pos relativ zu MCS"
    Rectangle (16,430 95x19), "Translation"
END_VISUALIZATION

// Device/Application/VISU_Konfig
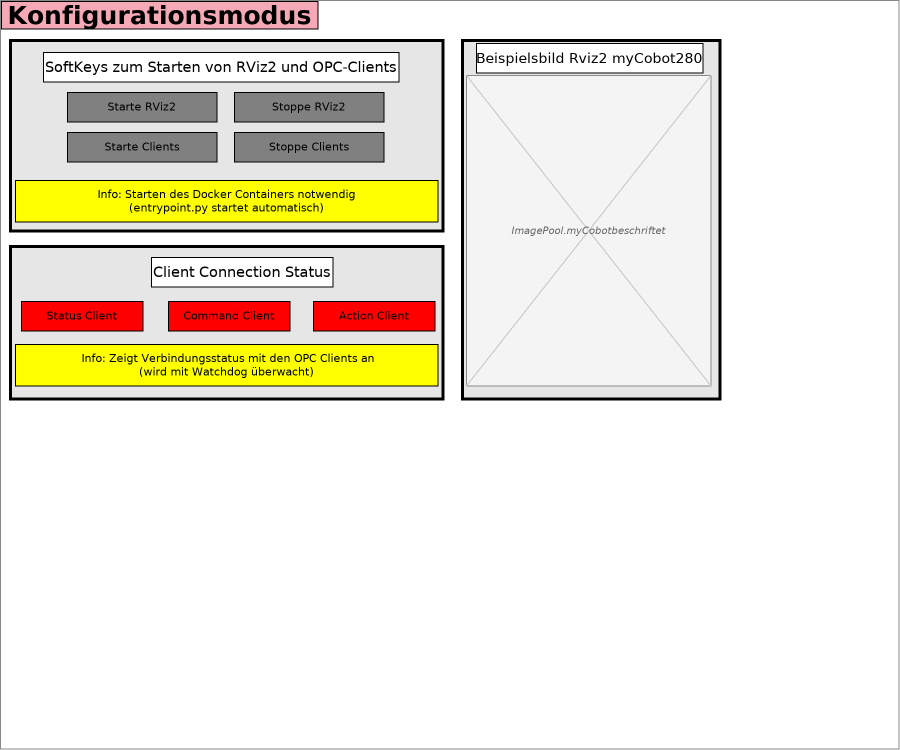
VISUALIZATION VISU_Konfig  // 900x750
    Rectangle (1,1 317x28), "Konfigurationsmodus"
    Rectangle (461,39 260x361)
    Rectangle (9,39 435x193)
    Rectangle (67,92 150x30), "Starte RViz2"
        toggle GVL_OPCUA.Start_RViz2
        OnMouseClick: execute { GVL_OPCUA.Stop_RViz2 := FALSE; }
    Rectangle (67,132 150x30), "Starte Clients"
        toggle GVL_OPCUA.Start_OPCClients
        OnMouseClick: execute { GVL_OPCUA.Stop_OPC_Clients := False; }
    Rectangle (234,132 150x30), "Stoppe Clients"
        toggle GVL_OPCUA.Stop_OPC_Clients
        OnMouseClick: execute { GVL_OPCUA.Start_OPCClients := False; }
    Rectangle (234,92 150x30), "Stoppe RViz2"
        toggle GVL_OPCUA.Stop_RViz2
        OnMouseClick: execute { GVL_OPCUA.Start_RViz2 := FALSE; }
    Image (466,75 245x311), image: ImagePool.myCobotbeschriftet
    Rectangle (476,43 227x30), "Beispielsbild Rviz2 myCobot280"
    Rectangle (43,52 356x30), "SoftKeys zum Starten von RViz2 und OPC-Clients"
    Rectangle (15,180 423x42), "Info: Starten des Docker Containers notwendig (entrypoint.py startet automatisch)"
    Rectangle (9,245 435x155)
    Rectangle (151,257 182x30), "Client Connection Status"
    Rectangle (21,301 122x30), "Status Client", colour toggle: MAIN_PRG.RobotStatus.client_connected
    Rectangle (313,301 122x30), "Action Client", colour toggle: MAIN_PRG.RobotAction.client_connected
    Rectangle (168,301 122x30), "Command Client", colour toggle: MAIN_PRG.RobotCommand.client_connected
    Rectangle (15,344 423x42), "Info: Zeigt Verbindungsstatus mit den OPC Clients an (wird mit Watchdog überwacht)"
END_VISUALIZATION

// Device/Application/VISU_Schrittkette
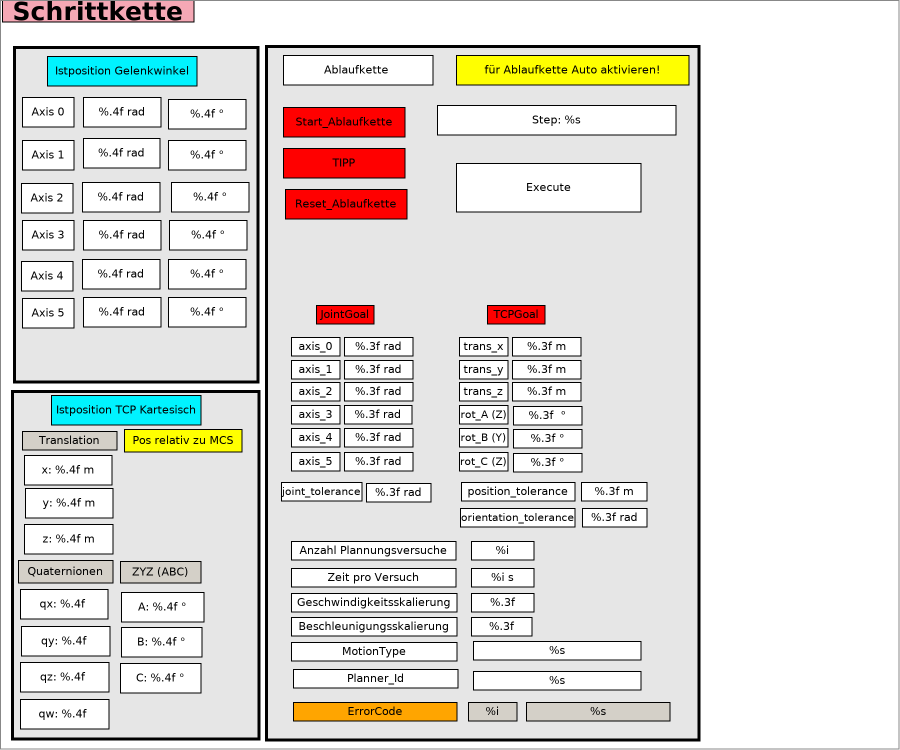
VISUALIZATION VISU_Schrittkette  // 900x750
    Rectangle (265,45 435x696)
    Rectangle (283,55 150x30), "Ablaufkette"
    Rectangle (283,148 122x30), "TIPP", colour toggle: MAIN_PRG.RobotStatus.client_connected
        tap GVL_OPCUA.TIPP
    Rectangle (283,107 122x30), "Start_Ablaufkette", colour toggle: MAIN_PRG.RobotStatus.client_connected
        tap GVL_OPCUA.Start_Ablaufkette
    Rectangle (437,105 239x30), "Step: %s", text variable: Ablaufkette.SFCCurrentStep
    Rectangle (456,55 233x30), "für Ablaufkette Auto aktivieren!"
    Rectangle (285,189 122x30), "Reset_Ablaufkette", colour toggle: MAIN_PRG.RobotStatus.client_connected
        tap GVL_OPCUA.Reset_Ablaufkette
    Rectangle (456,163 185x49), "Execute"
        tap GVL_OPCUA.Execute
    Rectangle (2,0 192x22), "Schrittkette"
    Rectangle (291,337 49x19), "axis_0"
    Rectangle (291,360 49x19), "axis_1"
    Rectangle (291,382 49x19), "axis_2"
    Rectangle (291,405 49x19), "axis_3"
    Rectangle (291,428 49x19), "axis_4"
    Rectangle (291,452 49x19), "axis_5"
    Rectangle (344,337 69x19), "%.3f rad", text variable: MAIN_PRG.RobotAction.axis_0
        OnMouseClick: write the text variable via Default
    Rectangle (344,360 69x19), "%.3f rad", text variable: MAIN_PRG.RobotAction.axis_1
        OnMouseClick: write the text variable via Default
    Rectangle (344,382 69x19), "%.3f rad", text variable: MAIN_PRG.RobotAction.axis_2
        OnMouseClick: write the text variable via Default
    Rectangle (344,405 68x19), "%.3f rad", text variable: MAIN_PRG.RobotAction.axis_3
        OnMouseClick: write the text variable via Default
    Rectangle (344,428 69x19), "%.3f rad", text variable: MAIN_PRG.RobotAction.axis_4
        OnMouseClick: write the text variable via Default
    Rectangle (344,452 69x19), "%.3f rad", text variable: MAIN_PRG.RobotAction.axis_5
        OnMouseClick: write the text variable via Default
    Rectangle (459,337 49x19), "trans_x"
    Rectangle (459,360 49x19), "trans_y"
    Rectangle (459,382 49x19), "trans_z"
    Rectangle (512,337 69x19), "%.3f m", text variable: MAIN_PRG.RobotAction.trans_x
        OnMouseClick: write the text variable via Default
    Rectangle (512,360 69x19), "%.3f m", text variable: MAIN_PRG.RobotAction.trans_y
        OnMouseClick: write the text variable via Default
    Rectangle (512,382 69x19), "%.3f m", text variable: MAIN_PRG.RobotAction.trans_z
        OnMouseClick: write the text variable via Default
    Rectangle (316,305 58x19), "JointGoal", colour toggle: MAIN_PRG.RobotAction.Joint_Goal
        toggle MAIN_PRG.RobotAction.Joint_Goal
    Rectangle (487,305 58x19), "TCPGoal", colour toggle: MAIN_PRG.RobotAction.TCP_Goal
        toggle MAIN_PRG.RobotAction.TCP_Goal
    Rectangle (291,541 165x19), "Anzahl Plannungsversuche"
    Rectangle (291,568 165x19), "Zeit pro Versuch"
    Rectangle (291,593 166x19), "Geschwindigkeitsskalierung"
    Rectangle (291,617 166x19), "Beschleunigungsskalierung"
    Rectangle (461,482 114x19), "position_tolerance"
    Rectangle (460,508 115x19), "orientation_tolerance"
    Rectangle (471,541 63x19), "%i", text variable: MAIN_PRG.RobotAction.num_planning_attempts
        OnMouseClick: write the text variable via Default
    Rectangle (471,568 63x19), "%i s", text variable: MAIN_PRG.RobotAction.allowed_planning_time
        OnMouseClick: write the text variable via Default
    Rectangle (471,593 63x19), "%.3f", text variable: MAIN_PRG.RobotAction.max_velocity_scaling
        OnMouseClick: write the text variable via Default
    Rectangle (471,617 61x19), "%.3f", text variable: MAIN_PRG.RobotAction.max_acceleration_scaling
        OnMouseClick: write the text variable via Default
    Rectangle (581,482 66x19), "%.3f m", text variable: MAIN_PRG.RobotAction.position_tolerance
        OnMouseClick: write the text variable via Default
    Rectangle (582,508 65x19), "%.3f rad", text variable: MAIN_PRG.RobotAction.orientation_tolerance
        OnMouseClick: write the text variable via Default
    Rectangle (291,642 166x19), "MotionType"
    Rectangle (293,669 165x19), "Planner_Id"
    Rectangle (293,702 164x19), "ErrorCode"
    Rectangle (468,702 49x19), "%i", text variable: MAIN_PRG.RobotAction.error_code
    Rectangle (473,641 168x19), "%s", text variable: MAIN_PRG.RobotAction.Motion_Type
        OnMouseClick: write the text variable via Default
    Rectangle (473,671 168x19), "%s", text variable: MAIN_PRG.RobotAction.Planner_ID
        OnMouseClick: write the text variable via Default
    Rectangle (526,702 144x19), "%s", text variable: MAIN_PRG.Status_Error_Codes_Action
    Rectangle (459,405 49x19), "rot_A (Z)"
    Rectangle (459,428 49x19), "rot_B (Y)"
    Rectangle (459,452 49x19), "rot_C (Z)"
    Rectangle (513,406 69x19), "%.3f °", text variable: GVL_OPCUA.rot_A
        OnMouseClick: write the text variable via Default
    Rectangle (513,429 69x19), "%.3f °", text variable: GVL_OPCUA.rot_B
        OnMouseClick: write the text variable via Default
    Rectangle (513,453 69x19), "%.3f °", text variable: GVL_OPCUA.rot_C
        OnMouseClick: write the text variable via Default
    Rectangle (366,483 65x19), "%.3f rad", text variable: MAIN_PRG.RobotAction.joint_tolerance
        OnMouseClick: write the text variable via Default
    Rectangle (281,482 81x19), "joint_tolerance"
    Rectangle (11,390 249x350)
    Rectangle (13,46 246x337)
    Rectangle (47,56 150x30), "Istposition Gelenkwinkel"
    Rectangle (51,395 150x30), "Istposition TCP Kartesisch"
    Rectangle (24,455 88x30), "x: %.4f m", text variable: GVL_OPCUA.RobotStatus.Ist_Pos_TCP.trans_x
    Rectangle (25,488 88x30), "y: %.4f m", text variable: GVL_OPCUA.RobotStatus.Ist_Pos_TCP.trans_y
    Rectangle (24,524 89x30), "z: %.4f m", text variable: GVL_OPCUA.RobotStatus.Ist_Pos_TCP.trans_z
    Rectangle (20,589 88x30), "qx: %.4f", text variable: GVL_OPCUA.RobotStatus.Ist_Pos_TCP.rot_x
    Rectangle (21,626 89x30), "qy: %.4f", text variable: GVL_OPCUA.RobotStatus.Ist_Pos_TCP.rot_y
    Rectangle (20,662 89x30), "qz: %.4f", text variable: GVL_OPCUA.RobotStatus.Ist_Pos_TCP.rot_z
    Rectangle (20,699 89x30), "qw: %.4f", text variable: GVL_OPCUA.RobotStatus.Ist_Pos_TCP.rot_w
    Rectangle (83,97 78x30), "%.4f rad", text variable: GVL_OPCUA.RobotStatus.Ist_Pos_Axis.axis_0
    Rectangle (83,138 77x30), "%.4f rad", text variable: GVL_OPCUA.RobotStatus.Ist_Pos_Axis.axis_1
    Rectangle (82,182 78x30), "%.4f rad", text variable: GVL_OPCUA.RobotStatus.Ist_Pos_Axis.axis_2
    Rectangle (83,220 78x30), "%.4f rad", text variable: GVL_OPCUA.RobotStatus.Ist_Pos_Axis.axis_3
    Rectangle (82,259 78x30), "%.4f rad", text variable: GVL_OPCUA.RobotStatus.Ist_Pos_Axis.axis_4
    Rectangle (83,297 78x30), "%.4f rad", text variable: GVL_OPCUA.RobotStatus.Ist_Pos_Axis.axis_5
    Rectangle (168,99 78x30), "%.4f °", text variable: GVL_OPCUA.RobotStatus.Ist_Pos_Axis.axis_0 *(180.0/GVL_OPCUA.PI)
    Rectangle (168,140 78x30), "%.4f °", text variable: GVL_OPCUA.RobotStatus.Ist_Pos_Axis.axis_1 *(180.0/GVL_OPCUA.PI)
    Rectangle (171,182 78x30), "%.4f °", text variable: GVL_OPCUA.RobotStatus.Ist_Pos_Axis.axis_2 *(180.0/GVL_OPCUA.PI)
    Rectangle (169,220 78x30), "%.4f °", text variable: GVL_OPCUA.RobotStatus.Ist_Pos_Axis.axis_3 *(180.0/GVL_OPCUA.PI)
    Rectangle (168,259 78x30), "%.4f °", text variable: GVL_OPCUA.RobotStatus.Ist_Pos_Axis.axis_4 *(180.0/GVL_OPCUA.PI)
    Rectangle (168,297 78x30), "%.4f °", text variable: GVL_OPCUA.RobotStatus.Ist_Pos_Axis.axis_5 *(180.0/GVL_OPCUA.PI)
    Rectangle (121,592 83x30), "A: %.4f °", text variable: MAIN_PRG.Status_Quat_to_ZYZ.euler.A
    Rectangle (121,627 81x30), "B: %.4f °", text variable: MAIN_PRG.Status_Quat_to_ZYZ.euler.B
    Rectangle (120,663 81x30), "C: %.4f °", text variable: MAIN_PRG.Status_Quat_to_ZYZ.euler.C
    Rectangle (120,561 81x22), "ZYZ (ABC)"
    Rectangle (18,560 95x23), "Quaternionen"
    Rectangle (22,97 52x30), "Axis 0"
    Rectangle (22,140 52x30), "Axis 1"
    Rectangle (21,183 52x30), "Axis 2"
    Rectangle (22,220 52x30), "Axis 3"
    Rectangle (21,261 52x30), "Axis 4"
    Rectangle (22,298 52x30), "Axis 5"
    RoundedRectangle (124,429 118x23), "Pos relativ zu MCS"
    Rectangle (22,431 95x19), "Translation"
END_VISUALIZATION
